           #System.OrderTable[#Chain_To_Chain_CurrentOrder].Status := #CANCELED_STATUS;
           #System.OrderTable[#Chain_To_Chain_CurrentOrder].CompleteTime := #CurrentTime;
           #Chain_To_Chain_CurrentOrder := 0;
           //#Cnv_Entry.Instruction.Execute := FALSE;
       END_IF;

       //Error
       IF (#Cnv_PopUp_2.Error OR #Cnv_PopUp_3.Error) THEN
           //#Cnv_Entry.Instruction.Execute := FALSE;
           //
           "Control_DB"."Carrousel_Order Table".Task_Data_Available := FALSE;//#System.OrderTable[#Chain_To_Chain_CurrentOrder].OPC_Control.Task_Data_Available; // Send the Task Data Available from WCS 
           "Control_DB"."Carrousel_Order Table".Task_Type := 0; //  Send the Task Type - Chain to Chain Conveyor = Task Type = 7
           "Control_DB"."Carrousel_Order Table".Task_ID := 0; // Send the Task ID number;
           "Control_DB"."Carrousel_Order Table".Task_Metadata := ''; // Send the Task Metadata Unique identifier
           "Control_DB"."Carrousel_Order Table".Source_Location := 0; // Send the Source Location from the Conveyor
           "Control_DB"."Carrousel_Order Table".Destination_Location := 0; // Send the Destination Location to the Conveyor;

           #System.OrderTable[#Chain_To_Chain_CurrentOrder].ErrorID := (#Cnv_PopUp_2.Cnv_Errors.Error_Word_1
                                                                        OR #Cnv_PopUp_3.Cnv_Errors.Error_Word_1);

       END_IF;

       //MOVEMENT FINALIZED
       #Chain_To_ChainDoneRTrig(CLK := "Control_DB"."Carrousel_Order Table".Movement_Request_Complete);
       IF #Chain_To_ChainDoneRTrig.Q THEN

           "Control_DB"."Carrousel_Order Table".Task_Data_Available := FALSE;//#System.OrderTable[#Chain_To_Chain_CurrentOrder].OPC_Control.Task_Data_Available; // Send the Task Data Available from WCS 
           "Control_DB"."Carrousel_Order Table".Task_Type := 0; //  Send the Task Type - Chain to Chain Conveyor = Task Type = 7
           "Control_DB"."Carrousel_Order Table".Task_ID := 0; // Send the Task ID number;
           "Control_DB"."Carrousel_Order Table".Task_Metadata := ''; // Send the Task Metadata Unique identifier
           "Control_DB"."Carrousel_Order Table".Source_Location := 0; // Send the Source Location from the Conveyor
           "Control_DB"."Carrousel_Order Table".Destination_Location := 0; // Send the Destination Location to the Conveyor;


           #Chain_To_Chain_WatchdogStart := FALSE;
           #System.OrderTable[#Chain_To_Chain_CurrentOrder].Status := #COMPLETED_STATUS;
           #System.OrderTable[#Chain_To_Chain_CurrentOrder].CompleteTime := #CurrentTime;
           #Chain_To_Chain_CurrentOrder := 0;
       END_IF;
   END_REGION

   REGION Pop4 to Pick Station - Carousel Conveyors - Pop 4 to Pick Station
       IF #System.OrderTable[1].StepNo <> 0
           AND #System.OrderTable[1].Device = #POP4_TO_PICK_DEVICE
           AND #System.OrderTable[1].Status = #QUEUED_STATUS
           AND NOT (#Cnv_PopUp_4.Running OR #Cnv_PopUp_1.Running)
           AND NOT #System.Error
           AND NOT #Canceling
           AND #System.OrderTable[#Roller_To_Roller_CurrentOrder].Status <> #RUNNING_STATUS
           AND #System.OrderTable[#PickSt_To_Pop1_CurrentOrder].Status <> #RUNNING_STATUS

       THEN
           #Pop4_To_PickSt_CurrentOrder := 1;
       END_IF;
       IF #System.OrderTable[#Pop4_To_PickSt_CurrentOrder].StepNo <> 0
           AND #System.OrderTable[#Pop4_To_PickSt_CurrentOrder].Device = #POP4_TO_PICK_DEVICE
           AND #System.OrderTable[#Pop4_To_PickSt_CurrentOrder].Status = #QUEUED_STATUS
           AND NOT (#Cnv_PopUp_4.Running OR #Cnv_PopUp_1.Running)
           AND NOT #System.Error
           AND NOT #Canceling
           AND #System.OrderTable[#Roller_To_Roller_CurrentOrder].Status <> #RUNNING_STATUS
           AND #System.OrderTable[#PickSt_To_Pop1_CurrentOrder].Status <> #RUNNING_STATUS
       THEN
           //OPC Commands to Move Pallets - Carousel Conveyors
           // WCS => Order Table => OPC Ua Control Table

           "Control_DB"."Carrousel_Order Table".Task_Data_Available := TRUE;//#System.OrderTable[#Pop4_To_PickSt_CurrentOrder].OPC_Control.Task_Data_Available; // Send the Task Data Available from WCS 
           "Control_DB"."Carrousel_Order Table".Task_Type := #System.OrderTable[#Pop4_To_PickSt_CurrentOrder].OPC_Control.Task_Type; //  Send the Task Type - Pop4 to Pick Station Conveyor = Task Type = 8
           "Control_DB"."Carrousel_Order Table".Task_ID := #System.OrderTable[#Pop4_To_PickSt_CurrentOrder].OPC_Control.Task_ID; // Send the Task ID number;
           "Control_DB"."Carrousel_Order Table".Task_Metadata := #System.OrderTable[#Pop4_To_PickSt_CurrentOrder].OPC_Control.Task_Metadata; // Send the Task Metadata Unique identifier
           "Control_DB"."Carrousel_Order Table".Source_Location := #System.OrderTable[#Pop4_To_PickSt_CurrentOrder].OPC_Control.Source_Location; // Send the Source Location from the Conveyor
           "Control_DB"."Carrousel_Order Table".Destination_Location := #System.OrderTable[#Pop4_To_PickSt_CurrentOrder].OPC_Control.Destination_Location; // Send the Destination Location to the Conveyor;
           #Pop4_To_PickWatchdogStart := TRUE;



       END_IF;

       //RUNNING
       IF (#Cnv_PopUp_4.Running OR #Cnv_PopUp_1.Running) AND #System.Auto_Man THEN
           //#Cnv_Entry.Instruction.Execute := FALSE;
           #System.OrderTable[#Pop4_To_PickSt_CurrentOrder].Status := #RUNNING_STATUS;
       END_IF;

       //Cancel order
       IF #Canceling AND NOT (#Cnv_PopUp_4.Running OR #Cnv_PopUp_1.Running) AND #Pop4_To_PickSt_CurrentOrder <> 0 THEN
           #System.OrderTable[#Pop4_To_PickSt_CurrentOrder].Status := #CANCELED_STATUS;
           #System.OrderTable[#Pop4_To_PickSt_CurrentOrder].CompleteTime := #CurrentTime;
           #Pop4_To_PickSt_CurrentOrder := 0;

           "Control_DB"."Carrousel_Order Table".Task_Data_Available := FALSE;//#System.OrderTable[#Chain_To_Chain_CurrentOrder].OPC_Control.Task_Data_Available; // Send the Task Data Available from WCS 
           "Control_DB"."Carrousel_Order Table".Task_Type := 0; //  Send the Task Type - Chain to Chain Conveyor = Task Type = 7
           "Control_DB"."Carrousel_Order Table".Task_ID := 0; // Send the Task ID number;
           "Control_DB"."Carrousel_Order Table".Task_Metadata := ''; // Send the Task Metadata Unique identifier
           "Control_DB"."Carrousel_Order Table".Source_Location := 0; // Send the Source Location from the Conveyor
           "Control_DB"."Carrousel_Order Table".Destination_Location := 0; // Send the Destination Location to the Conveyor;

           //#Cnv_Entry.Instruction.Execute := FALSE;
       END_IF;

       //Error
       IF (#Cnv_PopUp_4.Error OR #Cnv_PopUp_1.Error) THEN
           //#Cnv_Entry.Instruction.Execute := FALSE;
           "Control_DB"."Carrousel_Order Table".Task_Data_Available := FALSE;//#System.OrderTable[#Chain_To_Chain_CurrentOrder].OPC_Control.Task_Data_Available; // Send the Task Data Available from WCS 
           "Control_DB"."Carrousel_Order Table".Task_Type := 0; //  Send the Task Type - Chain to Chain Conveyor = Task Type = 7
           "Control_DB"."Carrousel_Order Table".Task_ID := 0; // Send the Task ID number;
           "Control_DB"."Carrousel_Order Table".Task_Metadata := ''; // Send the Task Metadata Unique identifier
           "Control_DB"."Carrousel_Order Table".Source_Location := 0; // Send the Source Location from the Conveyor
           "Control_DB"."Carrousel_Order Table".Destination_Location := 0; // Send the Destination Location to the Conveyor;
           #System.OrderTable[#Pop4_To_PickSt_CurrentOrder].ErrorID := (#Cnv_PopUp_4.Cnv_Errors.Error_Word_1
           OR #Cnv_PopUp_1.Cnv_Errors.Error_Word_1);

       END_IF;

       //MOVEMENT FINALIZED
       #Pop4_To_PickSt_DoneRTrig(CLK := "Control_DB"."Carrousel_Order Table".Movement_Request_Complete);
       IF #Pop4_To_PickSt_DoneRTrig.Q THEN
           #Pop4_To_PickWatchdogStart := FALSE;

           "Control_DB"."Carrousel_Order Table".Task_Data_Available := FALSE;//#System.OrderTable[#Chain_To_Chain_CurrentOrder].OPC_Control.Task_Data_Available; // Send the Task Data Available from WCS 
           "Control_DB"."Carrousel_Order Table".Task_Type := 0; //  Send the Task Type - Chain to Chain Conveyor = Task Type = 7
           "Control_DB"."Carrousel_Order Table".Task_ID := 0; // Send the Task ID number;
           "Control_DB"."Carrousel_Order Table".Task_Metadata := ''; // Send the Task Metadata Unique identifier
           "Control_DB"."Carrousel_Order Table".Source_Location := 0; // Send the Source Location from the Conveyor
           "Control_DB"."Carrousel_Order Table".Destination_Location := 0; // Send the Destination Location to the Conveyor;

           #System.OrderTable[#Pop4_To_PickSt_CurrentOrder].Status := #COMPLETED_STATUS;
           #System.OrderTable[#Pop4_To_PickSt_CurrentOrder].CompleteTime := #CurrentTime;
           #Pop4_To_PickSt_CurrentOrder := 0;
       END_IF;
   END_REGION

   REGION Pick Station to Pop1 - Carousel Conveyors - Pick Station To Pop 1 
       IF #System.OrderTable[1].StepNo <> 0
           AND #System.OrderTable[1].Device = #PICK_TO_POP1_DEVICE
           AND #System.OrderTable[1].Status = #QUEUED_STATUS
           AND NOT (#Cnv_PopUp_1.Running)
           AND NOT #System.Error
           AND NOT #Canceling
           AND #System.OrderTable[#Roller_To_Roller_CurrentOrder].Status <> #RUNNING_STATUS
           AND #System.OrderTable[#Pop4_To_PickSt_CurrentOrder].Status <> #RUNNING_STATUS
       THEN
           #PickSt_To_Pop1_CurrentOrder := 1;
       END_IF;
       IF #System.OrderTable[#PickSt_To_Pop1_CurrentOrder].StepNo <> 0
           AND #System.OrderTable[#PickSt_To_Pop1_CurrentOrder].Device = #PICK_TO_POP1_DEVICE
           AND #System.OrderTable[#PickSt_To_Pop1_CurrentOrder].Status = #QUEUED_STATUS
           AND NOT (#Cnv_PopUp_1.Running)
           AND NOT #System.Error
           AND NOT #Canceling
           AND #System.OrderTable[#Roller_To_Roller_CurrentOrder].Status <> #RUNNING_STATUS
           AND #System.OrderTable[#Pop4_To_PickSt_CurrentOrder].Status <> #RUNNING_STATUS
       THEN
           //OPC Commands to Move Pallets - Carousel Conveyors
           // WCS => Order Table => OPC Ua Control Table

           "Control_DB"."Carrousel_Order Table".Task_Data_Available := TRUE;//#System.OrderTable[#PickSt_To_Pop1_CurrentOrder].OPC_Control.Task_Data_Available; // Send the Task Data Available from WCS 
           "Control_DB"."Carrousel_Order Table".Task_Type := #System.OrderTable[#PickSt_To_Pop1_CurrentOrder].OPC_Control.Task_Type; //  Send the Task Type - Roller to Roller Conveyor = Task Type = 6
           "Control_DB"."Carrousel_Order Table".Task_ID := #System.OrderTable[#PickSt_To_Pop1_CurrentOrder].OPC_Control.Task_ID; // Send the Task ID number;
           "Control_DB"."Carrousel_Order Table".Task_Metadata := #System.OrderTable[#PickSt_To_Pop1_CurrentOrder].OPC_Control.Task_Metadata; // Send the Task Metadata Unique identifier
           "Control_DB"."Carrousel_Order Table".Source_Location := #System.OrderTable[#PickSt_To_Pop1_CurrentOrder].OPC_Control.Source_Location; // Send the Source Location from the Conveyor
           "Control_DB"."Carrousel_Order Table".Destination_Location := #System.OrderTable[#PickSt_To_Pop1_CurrentOrder].OPC_Control.Destination_Location; // Send the Destination Location to the Conveyor;
           #PickSt_To_Pop1WatchdogStart := true;


       END_IF;

       //RUNNING
       IF (#Cnv_PopUp_1.Running) AND #System.Auto_Man THEN
           //#Cnv_Entry.Instruction.Execute := FALSE;
           #System.OrderTable[#PickSt_To_Pop1_CurrentOrder].Status := #RUNNING_STATUS;
       END_IF;

       //Cancel order
       IF #Canceling AND NOT (#Cnv_PopUp_1.Running) AND #PickSt_To_Pop1_CurrentOrder <> 0 THEN
           #System.OrderTable[#PickSt_To_Pop1_CurrentOrder].Status := #CANCELED_STATUS;
           #System.OrderTable[#PickSt_To_Pop1_CurrentOrder].CompleteTime := #CurrentTime;
           #PickSt_To_Pop1_CurrentOrder := 0;
           "Control_DB"."Carrousel_Order Table".Task_Data_Available := FALSE;//#System.OrderTable[#Chain_To_Chain_CurrentOrder].OPC_Control.Task_Data_Available; // Send the Task Data Available from WCS 
           "Control_DB"."Carrousel_Order Table".Task_Type := 0; //  Send the Task Type - Chain to Chain Conveyor = Task Type = 7
           "Control_DB"."Carrousel_Order Table".Task_ID := 0; // Send the Task ID number;
           "Control_DB"."Carrousel_Order Table".Task_Metadata := ''; // Send the Task Metadata Unique identifier
           "Control_DB"."Carrousel_Order Table".Source_Location := 0; // Send the Source Location from the Conveyor
           "Control_DB"."Carrousel_Order Table".Destination_Location := 0; // Send the Destination Location to the Conveyor;
           //#Cnv_Entry.Instruction.Execute := FALSE;
       END_IF;

       //Error
       IF (#Cnv_PopUp_2.Error OR #Cnv_PopUp_3.Error) THEN
           //#Cnv_Entry.Instruction.Execute := FALSE;
           "Control_DB"."Carrousel_Order Table".Task_Data_Available := FALSE;//#System.OrderTable[#Chain_To_Chain_CurrentOrder].OPC_Control.Task_Data_Available; // Send the Task Data Available from WCS 
           "Control_DB"."Carrousel_Order Table".Task_Type := 0; //  Send the Task Type - Chain to Chain Conveyor = Task Type = 7
           "Control_DB"."Carrousel_Order Table".Task_ID := 0; // Send the Task ID number;
           "Control_DB"."Carrousel_Order Table".Task_Metadata := ''; // Send the Task Metadata Unique identifier
           "Control_DB"."Carrousel_Order Table".Source_Location := 0; // Send the Source Location from the Conveyor
           "Control_DB"."Carrousel_Order Table".Destination_Location := 0; // Send the Destination Location to the Conveyor;
           #System.OrderTable[#PickSt_To_Pop1_CurrentOrder].ErrorID := (#Cnv_PopUp_2.Cnv_Errors.Error_Word_1
           OR #Cnv_PopUp_3.Cnv_Errors.Error_Word_1);

       END_IF;

       //MOVEMENT FINALIZED
       #PickSt_To_Pop1_DoneRTrig(CLK := "Control_DB"."Carrousel_Order Table".Movement_Request_Complete);
       IF #PickSt_To_Pop1_DoneRTrig.Q THEN

           "Control_DB"."Carrousel_Order Table".Task_Data_Available := FALSE;//#System.OrderTable[#Chain_To_Chain_CurrentOrder].OPC_Control.Task_Data_Available; // Send the Task Data Available from WCS 
           "Control_DB"."Carrousel_Order Table".Task_Type := 0; //  Send the Task Type - Chain to Chain Conveyor = Task Type = 7
           "Control_DB"."Carrousel_Order Table".Task_ID := 0; // Send the Task ID number;
           "Control_DB"."Carrousel_Order Table".Task_Metadata := ''; // Send the Task Metadata Unique identifier
           "Control_DB"."Carrousel_Order Table".Source_Location := 0; // Send the Source Location from the Conveyor
           "Control_DB"."Carrousel_Order Table".Destination_Location := 0; // Send the Destination Location to the Conveyor;

           #PickSt_To_Pop1WatchdogStart := FALSE;
           #System.OrderTable[#PickSt_To_Pop1_CurrentOrder].Status := #COMPLETED_STATUS;
           #System.OrderTable[#PickSt_To_Pop1_CurrentOrder].CompleteTime := #CurrentTime;
           #PickSt_To_Pop1_CurrentOrder := 0;
       END_IF;
   END_REGION

   REGION Weigh Station - Carousel Conveyors 
       IF #System.OrderTable[1].StepNo <> 0
           AND #System.OrderTable[1].Device = #WEIGH_STATION_DEVICE
           AND #System.OrderTable[1].Status = #QUEUED_STATUS
           AND NOT ("Control_DB"."Weighing Station".Running)
           AND NOT #System.Error
           AND NOT #Canceling
       THEN
           #WeighingStation_CurrentOrder := 1;
       END_IF;
       IF #System.OrderTable[#WeighingStation_CurrentOrder].StepNo <> 0
           AND #System.OrderTable[#WeighingStation_CurrentOrder].Device = #WEIGH_STATION_DEVICE
           AND #System.OrderTable[#WeighingStation_CurrentOrder].Status = #QUEUED_STATUS
           AND NOT ("Control_DB"."Weighing Station".Running)
           AND NOT #System.Error
           AND NOT #Canceling
       THEN
           //OPC Commands to Move Pallets - Carousel Conveyors
           // WCS => Order Table => OPC Ua Control Table


           "Control_DB"."Carrousel_Order Table".Task_Data_Available := TRUE;//#System.OrderTable[#WeighingStation_CurrentOrder].OPC_Control.Task_Data_Available; // Send the Task Data Available from WCS 
           "Control_DB"."Carrousel_Order Table".Task_Type := #System.OrderTable[#WeighingStation_CurrentOrder].OPC_Control.Task_Type; //  Send the Task Type - Start Weigh Station = Task Type = 10
           "Control_DB"."Carrousel_Order Table".Task_ID := #System.OrderTable[#WeighingStation_CurrentOrder].OPC_Control.Task_ID; // Send the Task ID number;
           "Control_DB"."Carrousel_Order Table".Task_Metadata := #System.OrderTable[#WeighingStation_CurrentOrder].OPC_Control.Task_Metadata; // Send the Task Metadata Unique identifier
           #WeighingStation_WatchdogStart := true;


       END_IF;

       //RUNNING
       IF ("Control_DB"."Weighing Station".Running) AND #System.Auto_Man THEN
           //#Cnv_Entry.Instruction.Execute := FALSE;
           #System.OrderTable[#WeighingStation_CurrentOrder].Status := #RUNNING_STATUS;

       END_IF;

       //Cancel order
       IF #Canceling AND NOT ("Control_DB"."Weighing Station".Running) AND #WeighingStation_CurrentOrder <> 0 THEN
           #System.OrderTable[#WeighingStation_CurrentOrder].Status := #CANCELED_STATUS;
           #System.OrderTable[#WeighingStation_CurrentOrder].CompleteTime := #CurrentTime;
           #WeighingStation_CurrentOrder := 0;
           //#Cnv_Entry.Instruction.Execute := FALSE;
           "Control_DB"."Carrousel_Order Table".Task_Data_Available := FALSE;//#System.OrderTable[#WeighingStation_CurrentOrder].OPC_Control.Task_Data_Available; // Send the Task Data Available from WCS 
           "Control_DB"."Carrousel_Order Table".Task_Type := 0; //  Send the Task Type - Start Weigh Station = Task Type = 10
           "Control_DB"."Carrousel_Order Table".Task_ID := 0; // Send the Task ID number;
           "Control_DB"."Carrousel_Order Table".Task_Metadata := ''; // Send the Task Metadata Unique identifier
       END_IF;
     (*  
       //Error
       IF (#WeighingStation. OR #Cnv_PopUp_3.Error) THEN
           //#Cnv_Entry.Instruction.Execute := FALSE;

           #System.OrderTable[#WeighingStation_CurrentOrder].ErrorID := (#Cnv_PopUp_2.Cnv_Errors.Error_Word_1
         OR #Cnv_PopUp_3.Cnv_Errors.Error_Word_1);

       END_IF;
      *) 
       //MOVEMENT FINALIZED
       #WeighingStationDoneRTrig(CLK := "Control_DB"."Weighing Station".Done);
       IF #WeighingStationDoneRTrig.Q THEN
           #WeighingStation_WatchdogStart := FALSE;
           #System.OrderTable[#WeighingStation_CurrentOrder].Status := #COMPLETED_STATUS;
           #System.OrderTable[#WeighingStation_CurrentOrder].CompleteTime := #CurrentTime;
           #WeighingStation_CurrentOrder := 0;

           "Control_DB"."Carrousel_Order Table".Task_Data_Available := FALSE;//#System.OrderTable[#WeighingStation_CurrentOrder].OPC_Control.Task_Data_Available; // Send the Task Data Available from WCS 
           "Control_DB"."Carrousel_Order Table".Task_Type := 0; //  Send the Task Type - Start Weigh Station = Task Type = 10
           "Control_DB"."Carrousel_Order Table".Task_ID := 0; // Send the Task ID number;
           "Control_DB"."Carrousel_Order Table".Task_Metadata := ''; // Send the Task Metadata Unique identifier
       END_IF;
   END_REGION
   (*
   REGION Profile Station - Carousel Conveyors 
       IF #System.OrderTable[1].StepNo <> 0
           AND #System.OrderTable[1].Device = #PROFILE_STATION_DEVICE
           AND #System.OrderTable[1].Status = #QUEUED_STATUS
           AND NOT ("Control_DB"."Profiling Station".Running)
           AND NOT #System.Error
           AND NOT #Canceling
       THEN
           #ProfileStation_CurrentOrder := 1;
       END_IF;
       IF #System.OrderTable[#ProfileStation_CurrentOrder].StepNo <> 0
           AND #System.OrderTable[#ProfileStation_CurrentOrder].Device = #PROFILE_STATION_DEVICE
           AND #System.OrderTable[#ProfileStation_CurrentOrder].Status = #QUEUED_STATUS
           AND NOT ("Control_DB"."Profiling Station".Running)
           AND NOT #System.Error
           AND NOT #Canceling
       THEN
           //OPC Commands to Move Pallets - Carousel Conveyors
           // WCS => Order Table => OPC Ua Control Table

           "Control_DB"."Carrousel_Order Table".Task_Data_Available := TRUE;//#System.OrderTable[#ProfileStation_CurrentOrder].OPC_Control.Task_Data_Available; // Send the Task Data Available from WCS 
           "Control_DB"."Carrousel_Order Table".Task_Type := #System.OrderTable[#ProfileStation_CurrentOrder].OPC_Control.Task_Type; //  Send the Task Type - Start Weigh Station = Task Type = 10
           "Control_DB"."Carrousel_Order Table".Task_ID := #System.OrderTable[#ProfileStation_CurrentOrder].OPC_Control.Task_ID; // Send the Task ID number;
           "Control_DB"."Carrousel_Order Table".Task_Metadata := #System.OrderTable[#ProfileStation_CurrentOrder].OPC_Control.Task_Metadata; // Send the Task Metadata Unique identifier
           #ProfileStation_WatchdogStart := true;


       END_IF;

       //RUNNING
       IF ("Control_DB"."Profiling Station".Running) AND #System.Auto_Man THEN
           //#Cnv_Entry.Instruction.Execute := FALSE;
           #System.OrderTable[#ProfileStation_CurrentOrder].Status := #RUNNING_STATUS;

           "Control_DB"."Carrousel_Order Table".Task_Data_Available := FALSE;//#System.OrderTable[#ProfileStation_CurrentOrder].OPC_Control.Task_Data_Available; // Send the Task Data Available from WCS 
           "Control_DB"."Carrousel_Order Table".Task_Type := 0; //  Send the Task Type - Start Weigh Station = Task Type = 10
           "Control_DB"."Carrousel_Order Table".Task_ID := 0; // Send the Task ID number;
           "Control_DB"."Carrousel_Order Table".Task_Metadata := ''; // Send the Task Metadata Unique identifier
           #ProfileStation_WatchdogStart := true;
       END_IF;

       //Cancel order
       IF #Canceling AND NOT ("Control_DB"."Profiling Station".Running) AND #ProfileStation_CurrentOrder <> 0 THEN
           #System.OrderTable[#ProfileStation_CurrentOrder].Status := #CANCELED_STATUS;
           #System.OrderTable[#ProfileStation_CurrentOrder].CompleteTime := #CurrentTime;
           #ProfileStation_CurrentOrder := 0;
           "Control_DB"."Carrousel_Order Table".Task_Data_Available := FALSE;//#System.OrderTable[#ProfileStation_CurrentOrder].OPC_Control.Task_Data_Available; // Send the Task Data Available from WCS 
           "Control_DB"."Carrousel_Order Table".Task_Type := 0; //  Send the Task Type - Start Weigh Station = Task Type = 10
           "Control_DB"."Carrousel_Order Table".Task_ID := 0; // Send the Task ID number;
           "Control_DB"."Carrousel_Order Table".Task_Metadata := ''; // Send the Task Metadata Unique identifier
           //#Cnv_Entry.Instruction.Execute := FALSE;
       END_IF;
       (*  
         //Error
         IF (#WeighingStation. OR #Cnv_PopUp_3.Error) THEN
             //#Cnv_Entry.Instruction.Execute := FALSE;

             #System.OrderTable[#WeighingStation_CurrentOrder].ErrorID := (#Cnv_PopUp_2.Cnv_Errors.Error_Word_1
           OR #Cnv_PopUp_3.Cnv_Errors.Error_Word_1);

         END_IF;
        *)
        //MOVEMENT FINALIZED
       #ProfileStationDoneRTrig(CLK := "Control_DB"."Profiling Station".Done);
       IF #ProfileStationDoneRTrig.Q THEN
            #ProfileStation_WatchdogStart := FALSE;
            #System.OrderTable[#ProfileStation_CurrentOrder].Status := #COMPLETED_STATUS;
            #System.OrderTable[#ProfileStation_CurrentOrder].CompleteTime := #CurrentTime;
            #ProfileStation_CurrentOrder := 0;
            "Control_DB"."Carrousel_Order Table".Task_Data_Available := FALSE;//#System.OrderTable[#ProfileStation_CurrentOrder].OPC_Control.Task_Data_Available; // Send the Task Data Available from WCS 
            "Control_DB"."Carrousel_Order Table".Task_Type := 0; //  Send the Task Type - Start Weigh Station = Task Type = 10
            "Control_DB"."Carrousel_Order Table".Task_ID := 0; // Send the Task ID number;
            "Control_DB"."Carrousel_Order Table".Task_Metadata := ''; // Send the Task Metadata Unique identifier
        END_IF;
    END_REGION
   *)
   REGION Max Running Order Number
       #MaxRunningOrderNo := MAX(IN1 := #Roller_To_Roller_CurrentOrder, IN2 := #Chain_To_Chain_CurrentOrder,
                                 IN3 := #Pop4_To_PickSt_CurrentOrder, IN4 := #PickSt_To_Pop1_CurrentOrder,
                                 IN5 := #WeighingStation_CurrentOrder, IN6 := #ProfileStation_CurrentOrder);
   END_REGION

   REGION Pause Orders
       #ErrorRTrig(CLK := #System.Error);
       #PauseRTrig(CLK := #System.PauseOrders OR NOT #System.Auto_Man);
       IF #ErrorRTrig.Q OR #PauseRTrig.Q THEN
           #System.PauseOrders := FALSE;
           #System.Paused := #MaxRunningOrderNo > 0;
           IF #System.Paused THEN
               FOR #i := 1 TO UDINT_TO_DINT(#MaxRunningOrderNo) DO
                   IF #System.OrderTable[#i].Status = '' THEN
                       EXIT;
                   ELSIF #System.OrderTable[#i].Status = #QUEUED_STATUS THEN
                       #System.OrderTable[#i].Status := #PAUSED_STATUS;
                   ELSIF #System.OrderTable[#i].Status = #RUNNING_STATUS AND NOT #System.Auto_Man THEN
                       #System.OrderTable[#i].Status := #CANCELED_STATUS;
                   END_IF;
               END_FOR;
           END_IF;
       END_IF;
       IF #System.Paused AND #MaxRunningOrderNo = 0 THEN
           #System.Paused := FALSE;
       END_IF;
   END_REGION

   REGION Cancel Orders
       #CancelRTrig(CLK := #System.CancelOrders);
       #WeighingStation.Cancel := #ProfileStation.Cancel := #CancelRTrig.Q;
       IF #CancelRTrig.Q THEN
           #Canceling := TRUE;
           #System.CancelOrders := FALSE;
           #System.Paused := FALSE;
           FOR #i := 1 TO UDINT_TO_DINT(#MaxRunningOrderNo) DO
               IF #System.OrderTable[#i].Status = '' THEN
                   CONTINUE;
               ELSIF #System.OrderTable[#i].Status = #PAUSED_STATUS
                   OR #System.OrderTable[#i].Status = #QUEUED_STATUS
               THEN
                   #System.OrderTable[#i].Status := #CANCELED_STATUS;
                   #System.OrderTable[#i].CompleteTime := #CurrentTime;
               ELSIF #System.OrderTable[#i].Status = #ERROR_STATUS
               THEN
                   #System.OrderTable[#i].Status := #ERROR_CANCELED_STATUS;
                   #System.OrderTable[#i].CompleteTime := #CurrentTime;
               END_IF;
           END_FOR;
           #System.CurrentOrder := 0;
       END_IF;
       IF #Canceling AND NOT (#Cnv_Entry.Running OR #Cnv_PopUp_1.Running OR #WeighingStation.Running OR #ProfileStation.Running
           OR #Cnv_PopUp_2.Running OR #Cnv_PopUp_3.Running OR #Cnv_PopUp_4.Running OR #Cnv_Exit.Running) THEN
           #Canceling := FALSE;
           #Roller_To_Roller_CurrentOrder := #Chain_To_Chain_CurrentOrder:= #PickSt_To_Pop1_CurrentOrder := #Pop4_To_PickSt_CurrentOrder := 0;
            #WeighingStation_CurrentOrder:= #ProfileStation_CurrentOrder := 0;
       END_IF;
   END_REGION

   REGION Resume Orders
       #ResumeRTrig(CLK := #System.ResumeOrders);
       IF #ResumeRTrig.Q THEN
           #System.ResumeOrders := FALSE;
           #System.CurrentOrder := #MaxRunningOrderNo;
           IF NOT #System.Error THEN
               #System.Paused := FALSE;
               FOR #i := 1 TO UDINT_TO_DINT(#MaxRunningOrderNo) DO
                   IF #System.OrderTable[#i].Status = '' THEN
                       EXIT;
                   ELSIF #System.OrderTable[#i].Status = #PAUSED_STATUS
                       OR #System.OrderTable[#i].Status = #ERROR_STATUS
                   THEN
                       #System.OrderTable[#i].Status := #QUEUED_STATUS;
                   END_IF;
               END_FOR;
           END_IF;

       END_IF;
   END_REGION

   REGION Order Handler
       IF #System.Running AND NOT #System.Error
           AND (#System.OrderTable[#System.CurrentOrder].Status = #COMPLETED_STATUS
           OR #System.OrderTable[#System.CurrentOrder].Status = #ERROR_STATUS
           OR #System.OrderTable[#System.CurrentOrder].Status = #ERROR_CANCELED_STATUS
           OR #System.OrderTable[#System.CurrentOrder].Sequence = 0)
       THEN
           IF #System.CurrentOrder > 0 THEN
               #System.CurrentOrder -= 1;
           ELSE
               #System.CurrentOrder := 0;
           END_IF;
       END_IF;
   END_REGION

   REGION Watchdogs
       //Watchdog Timers
       #PickSt_To_Pop1WatchdogTimer(IN := #PickSt_To_Pop1WatchdogStart,
                                    PT := UDINT_TO_TIME(#Watchdog.Pick_TO_Pop1 * 60000),
                                    Q => #System.Watchdog_TimeOut.Pick_TO_Pop1);
       #Roller_To_Roller_WatchdogTimer(IN := #Roller_To_Roller_WatchdogStart,
                                       PT := UDINT_TO_TIME(#Watchdog.Roller_TO_Roller * 60000),
                                       Q => #System.Watchdog_TimeOut.Roller_TO_Roller);
       #Chain_To_Chain_WatchdogTimer(IN := #Chain_To_Chain_WatchdogStart,
                                     PT := UDINT_TO_TIME(#Watchdog.Chain_TO_Chain * 60000),
                                     Q => #System.Watchdog_TimeOut.Chain_TO_Chain);
       #Pop4_To_PickWatchdogTimer(IN := #Pop4_To_PickWatchdogStart,
                                  PT := UDINT_TO_TIME(#Watchdog.Pop4_TO_Pick * 60000),
                                  Q => #System.Watchdog_TimeOut.Pop4_TO_Pick);
       #WeighingStation_WatchdogTimer(IN := #WeighingStation_WatchdogStart,
                                      PT := UDINT_TO_TIME(#Watchdog.Weigh_Station * 60000),
                                      Q => #System.Watchdog_TimeOut.Weigh_Station);
       #ProfileStation_WatchdogTimer(IN := #ProfileStation_WatchdogStart,
                                     PT := UDINT_TO_TIME(#Watchdog.Profile_Station * 60000),
                                     Q => #System.Watchdog_TimeOut.Profile_Station);

       //Reset  Watchdog Timers
       IF #System.Error OR #CancelRTrig.Q OR #PauseRTrig.Q OR "Reset_All" THEN
           #PickSt_To_Pop1WatchdogStart := FALSE;
           #Roller_To_Roller_WatchdogStart := FALSE;
           #Chain_To_Chain_WatchdogStart := FALSE;
           #Pop4_To_PickWatchdogStart := FALSE;
           #WeighingStation_WatchdogStart := FALSE;
           #ProfileStation_WatchdogStart := FALSE;

       END_IF;
   END_REGION

   REGION Reset Next Order Number
       IF #System.NextOrder > 1
           AND #CurrentDTL.HOUR = 0
           AND #CurrentDTL.MINUTE = 0
           AND #CurrentDTL.SECOND = 0
       THEN
           #System.NextOrder := 1;
       END_IF;

   END_REGION

   REGION #System Mode and State
       #System.Selected := #System_Selected; // System selected
       #System.Ready := NOT #System.Error AND #System.Selected;
       #System.Auto_Man := #AutoMan_Switch;
       #System.Running := #Cnv_Entry.Running OR #Cnv_PopUp_1.Running OR #WeighingStation.Running
       OR #ProfileStation.Running OR #Cnv_PopUp_3.Running OR #Cnv_PopUp_4.Running;

       #System.Error := #Cnv_Entry.Error OR #Cnv_PopUp_1.Error OR #Cnv_PopUp_2.Error OR #Cnv_PopUp_3.Error OR #Cnv_PopUp_4.Error
       OR #Cnv_Exit.Error ; (*Implement Weigh station error and Profile Station error*)
       #System.IDLE := NOT #System.Running AND NOT #System.Paused AND NOT #System.Error;
       IF #System.Running THEN
           #System.State := 1;
       ELSIF #System.Paused AND NOT #System.Error THEN
           #System.State := 2;
       ELSIF #System.Error THEN
           #System.State := 3;
       ELSE
           #System.State := 0;
       END_IF;
   END_REGION
END_FUNCTION_BLOCK

FUNCTION_BLOCK "PConveyor_1_FB_1"   // FB36, SCL
TITLE = Conveyor Instance FB
{ S7_Optimized_Access := 'TRUE' }
AUTHOR : Mertin Coetzee
VERSION : 0.1
// stored: AutoNumber true, IsIECCheckEnabled false, IsRetainMemResEnabled false, MemoryReserve 100, SetENOAutomatically false, UDAEnableTagReadback false
   VAR_INPUT
      Cnv_Settings : "PopUp_Cnv_Settings";
   END_VAR
   VAR_IN_OUT
      Cnv_Control : "PopUp_Cnv_Control";
      SinaSpeed_Roller : SinaSpeed;
      SinaSpeed_Chain : SinaSpeed;
      SinaSpeed_Lift : SinaSpeed;
   END_VAR
   VAR
      State : UInt;
      Timer_TC : TON_TIME;
      Timer_Transfer { S7_SetPoint := 'True'} : TON_TIME;
      Watchdog { S7_SetPoint := 'True'} : TON_TIME;
      Transfer_Direction { S7_SetPoint := 'True'} : String;
      MainSetpoint_Roller : Int;
      MainSetpoint_Chain : Int;
      MainSetpoint_Lift : Int;
      IEC_Timer_0_Instance_1 { S7_SetPoint := 'True'} : TON_TIME;
      R_TRIG_Instance { S7_SetPoint := 'True'} : R_TRIG;
   END_VAR
   VAR_TEMP
      Execute_Old : Bool;
      Stop_Old : Bool;
   END_VAR
BEGIN
   "R_TRIG_DB_13"(CLK := #Cnv_Control.Instruction.Execute AND NOT #Execute_Old);
   "R_TRIG_DB_14"(CLK := #Cnv_Control.Instruction.Stop AND NOT #Stop_Old);

   #Execute_Old := #Cnv_Control.Instruction.Execute;
   #Stop_Old := #Cnv_Control.Instruction.Stop;

   #Cnv_Control.Enabled := #Cnv_Control.Instruction.Enable;

   //MODES
   #Cnv_Control.Mode := #Cnv_Control.Instruction.Mode_Change;
   IF (#Cnv_Control.Mode = 1 OR #Cnv_Control.Mode = 5) AND NOT #Cnv_Control.Error THEN
       #State := 500;
   END_IF;

   #R_TRIG_Instance(CLK := #Cnv_Control.Mode = 3);
   IF #R_TRIG_Instance.Q THEN
       #State := 0;
   END_IF;

   (*
   TODO:
   01. Need to add statemachine watchdog - Done
   02. Extractor needs to be on same floor for pallet to be moved in manual passed Rbwd - Done
   03. Complete reset state - Done
   04. Add stop inputs - Done
   05. Need to add variable motor speed, manual needs to be slower. - Done
   06. Need to add cyclic error checking. For odd sensor combinations as well - Partially done
   07. Need to add Shuttle monitor - Done
   08. Need to add Task ID check and start bit check to outbound pallet move. Check direction of pallet movement based on connected Cnv.
   09. Need to add checks for wrong direction of travel - Done
   10. Add checks for unsafe conditions with Cnv_Inputs - Partially Done
   11. Define Error codes - DOne
   12. Add watchdof time to Cnv Settings - Done
   13. Add self-timeout on manual 
   14. For shuttle in place sensor checks take into account extractor floor and safety stopper state
   15. Confirm modes and states are correct (Semi-auto and maintenance as well)
   16. Add the correct transfer process for the logistex-spacemaker pallet handovers.

   Mode select is done via the HMI. Might add external mode select switches.

           Mode select mask:
           0: Disabled
           1: Manual
           2: Semi-Auto
           3: Auto
           4: Teach - N/A for Cnv
           5: Maintenance

   Device ID Format: XXYYZZ    
   XX = Device type   
       01   VTD
       10  Cnv_Front_of_VTD
       11  Cnv_Rear_of_VTD
       12  Cnv_On_Extractor
       20  Safety_Stop_Front_of_VTD
       21  Safety_Stop_Rear_of_VTD
   YY = Floor   
   ZZ = VTD Connected to    
   Example: 110203 Conveyor at the rear of VTD 3 on level 2

   Pallet Alignment
   0 = no alignment
   1 = center alignment
   2 = Left
   3 = Right

    Sensor order for the conveyor:
    Lfwd Lpd1 Lpd2
     []   []   []
    ##############################
    #        Pallet Flow         #
    #         ------->>          #
    #                            #
    #                            #
    ##############################
                     []   []   []
                    Rpd2 Rpd1 Rbwd      
   *)

   REGION Cyclic Checks    
       // Update the pallet type as the Cnv_Inputs are triggered.
       #Cnv_Control.Cnv_Occupied := "PopUp Conveyor 2 - Pallet present 3";

       // Update the Cnv_Control opbject
       #Cnv_Control.SM_State := #State;
       #Cnv_Control.Stopped := NOT #Cnv_Control.Running;
       IF #Cnv_Control.Instruction.Inbound_Ready OR #Cnv_Control.Instruction.Outbound_Ready THEN
           #Cnv_Control.Ready_For_Task := TRUE;
       ELSE
           #Cnv_Control.Ready_For_Task := FALSE;
       END_IF;
   END_REGION

   REGION Auto/Semi auto mode
       CASE #State OF
           0: //Initialization
               #Cnv_Control.Instruction.Transfer_Complete := 0;
               #Cnv_Control.Instruction.Transfer_in_Progress := FALSE;
               #Cnv_Control.Running := FALSE;
               #Cnv_Control.Roller_Motor.Forward := FALSE;
               #Cnv_Control.Roller_Motor.Reverse := FALSE;
               #Cnv_Control.Roller_Motor.Speed := 0;
               #Cnv_Control.Chain_Motor.Forward := FALSE;
               #Cnv_Control.Chain_Motor.Reverse := FALSE;
               #Cnv_Control.Chain_Motor.Speed := 0;
               #Cnv_Control.Lift_Motor.Forward := FALSE;
               #Cnv_Control.Lift_Motor.Reverse := FALSE;
               #Cnv_Control.Lift_Motor.Speed := 0;
               #Transfer_Direction := '';
               #Timer_Transfer(IN := FALSE,
                               PT := T#0ms);
               IF #Cnv_Control.Enabled AND (#Cnv_Control.Mode = 3 OR #Cnv_Control.Mode = 2) AND #Cnv_Control.Error = 0 THEN
                   #State := 10;
               END_IF;

           10: //Standby - Conveyor ready to receive instruction
               IF ("R_TRIG_DB_13".Q OR #Cnv_Control.Instruction.Start_Transfer) THEN
                   //Inbound Transfer
                   IF #Cnv_Control.Instruction.Inbound_Ready AND NOT #Cnv_Control.Running AND #Cnv_Control.Error = 0 THEN
                       //Check transfer ID FROM Inbound conveyor
                       IF  #Cnv_Control.Inputs."Lift Up" THEN
                           #Cnv_Control.Done := FALSE;
                           #Cnv_Control.Instruction.Transfer_in_Progress := TRUE;
                           #Cnv_Control.Current_Task_ID := #Cnv_Control.Instruction.Task_ID;
                           #State := 20;// Roller Running (Popup Up)
                       ELSIF "Pick Station" AND
                           #Cnv_Control.Inputs."Lift Down" (*AND "Control_DB".PopUp_Cnv[4].Inputs."Lift Down"*) THEN //TO pick station
                           #Cnv_Control.Done := FALSE;
                           #Cnv_Control.Instruction.Transfer_in_Progress := TRUE;
                           #Cnv_Control.Current_Task_ID := #Cnv_Control.Instruction.Task_ID;
                           #State := 30;// Chain Running (Popup Down) 
                       ELSIF NOT "Pick Station" (*AND "Control_DB".PopUp_Cnv[4].Inputs."Lift Down"*) THEN //FROM pick station
                           #Cnv_Control.Done := FALSE;
                           #Cnv_Control.Instruction.Transfer_in_Progress := TRUE;
                           #Cnv_Control.Current_Task_ID := #Cnv_Control.Instruction.Task_ID;
                           #State := 40;
                       ELSE
                           #Cnv_Control.Warning := 1; //Cannot transfer from that conveyor
                       END_IF;

                       //Outbound Transfer    
                   ELSIF #Cnv_Control.Instruction.Outbound_Ready AND NOT #Cnv_Control.Running AND #Cnv_Control.Error = 0 THEN
                       //Check transfer ID TO popup cpnveyor 2
                       IF #Cnv_Control.Inputs."Lift Up" AND "Control_DB".PopUp_Cnv[2].Inputs."Lift Up" THEN
                           #Cnv_Control.Done := FALSE;
                           #Cnv_Control.Instruction.Transfer_in_Progress := TRUE;
                           #Cnv_Control.Current_Task_ID := #Cnv_Control.Instruction.Task_ID;
                           #State := 50;
                       ELSE
                           #Cnv_Control.Warning := 1; //Cannot transfer TO that conveyor
                       END_IF;
                   ELSE
                       #Cnv_Control.Warning := 0;// No task that can be started, yet start bit has been made true.
                   END_IF;
               ELSIF #Cnv_Control.Instruction.Start_Transfer AND "Control_DB".VTD_Control.Current_Level <> 0 THEN
                   //Extractor not at the correct level
                   "Set_Bit_F"(Bit := 2,
                               Bit_Value := 1,
                               Var := #Cnv_Control.Cnv_Errors.Error_Word_3);
               END_IF;
               IF #Cnv_Control.Instruction.Lift_Up THEN
                   #Cnv_Control.Done := FALSE;
                   #State := 60; // Lift UP
               ELSIF #Cnv_Control.Instruction.Lift_Down THEN
                   #Cnv_Control.Done := FALSE;
                   #State := 70; // Lift Down
               END_IF;

           20: // Roller Running (Popup Up)
               #Cnv_Control.Running := TRUE;
               #Cnv_Control.Roller_Motor.Forward := TRUE;
               #Cnv_Control.Roller_Motor.Speed := #Cnv_Settings.Roller_Full_Speed;
               #Transfer_Direction := 'Foward';

               IF "R_TRIG_DB_14".Q OR "PopUp Conveyor 2 - Pallet present 3" THEN
                   #Cnv_Control.Done := TRUE;
                   #Cnv_Control.Roller_Motor.Forward := FALSE;
                   #Cnv_Control.Roller_Motor.Reverse := FALSE;
                   #Cnv_Control.Roller_Motor.Speed := 0;
                   #Transfer_Direction := '';
                   #State := 0;
               END_IF;

               //Monitor the transfer progress
               #Timer_Transfer(IN := "Control_DB".Inbound_Cnv.Running,
                               PT := UINT_TO_TIME(#Cnv_Settings.Roller_Transfer_Time) * 1000);
               //If the watchdog bites, kill the process
               IF #Timer_Transfer.Q THEN //14:1 Transfer timed out
                   "Set_Bit_F"(Bit := 3,
                               Bit_Value := 1,
                               Var := #Cnv_Control.Cnv_Errors.Error_Word_2);
               END_IF;

           30: // Chain Running (Popup Down)
               #Cnv_Control.Running := TRUE;
               #Cnv_Control.Chain_Motor.Forward := TRUE;
               #Cnv_Control.Chain_Motor.Speed := #Cnv_Settings.Chain_Full_Speed;
               #Transfer_Direction := 'Foward';

               IF "R_TRIG_DB_14".Q OR NOT "Pick Station" THEN
                   #Cnv_Control.Done := TRUE;
                   #Cnv_Control.Chain_Motor.Forward := FALSE;
                   #Cnv_Control.Chain_Motor.Reverse := FALSE;
                   #Cnv_Control.Chain_Motor.Speed := 0;
                   #Transfer_Direction := '';
                   #State := 0;
               END_IF;

               //Monitor the transfer progress
               #Timer_Transfer(IN := "LighGuard_Cut-Off Path 01",
                               PT := UINT_TO_TIME(#Cnv_Settings.Chain_Transfer_Time) * 1000);
               //If the watchdog bites, kill the process
               IF #Timer_Transfer.Q THEN //14:1 Transfer timed out
                   "Set_Bit_F"(Bit := 3,
                               Bit_Value := 1,
                               Var := #Cnv_Control.Cnv_Errors.Error_Word_2);
               END_IF;

           40: // Chain Running (Popup Down)
               #Cnv_Control.Running := TRUE;
               #Cnv_Control.Chain_Motor.Forward := TRUE;
               #Cnv_Control.Chain_Motor.Speed := #Cnv_Settings.Chain_Full_Speed;
               #Transfer_Direction := 'Foward';

               IF "R_TRIG_DB_14".Q OR "PopUp Conveyor 1 - Pallet sensor" THEN
                   #Cnv_Control.Done := TRUE;
                   #Cnv_Control.Chain_Motor.Forward := FALSE;
                   #Cnv_Control.Chain_Motor.Reverse := FALSE;
                   #Cnv_Control.Chain_Motor.Speed := 0;
                   #Transfer_Direction := '';
                   #State := 0;
               END_IF;

               //Monitor the transfer progress
               #Timer_Transfer(IN := "LighGuard_Cut-Off Path 01",
                               PT := UINT_TO_TIME(#Cnv_Settings.Chain_Transfer_Time) * 1000);
               //If the watchdog bites, kill the process
               IF #Timer_Transfer.Q THEN //14:1 Transfer timed out
                   "Set_Bit_F"(Bit := 3,
                               Bit_Value := 1,
                               Var := #Cnv_Control.Cnv_Errors.Error_Word_2);
               END_IF;

           50: // Roller Running (Popup Up)
               IF "Control_DB".PopUp_Cnv[2].Roller_Motor.Status.%X0 THEN//Is running
                   #Cnv_Control.Running := TRUE;
                   #Cnv_Control.Roller_Motor.Forward := TRUE;
                   #Cnv_Control.Roller_Motor.Speed := #Cnv_Settings.Roller_Full_Speed;
                   #Transfer_Direction := 'Foward';
               END_IF;

               IF "R_TRIG_DB_14".Q OR "PopUp Conveyor 2 - Pallet present 4" THEN
                   #Cnv_Control.Done := TRUE;
                   #Cnv_Control.Roller_Motor.Forward := FALSE;
                   #Cnv_Control.Roller_Motor.Reverse := FALSE;
                   #Cnv_Control.Roller_Motor.Speed := 0;
                   #Transfer_Direction := '';
                   #State := 0;
               END_IF;

               //Monitor the transfer progress
               #Timer_Transfer(IN := TRUE,
                               PT := UINT_TO_TIME(#Cnv_Settings.Roller_Transfer_Time) * 1000);
               //If the watchdog bites, kill the process
               IF #Timer_Transfer.Q THEN //14:1 Transfer timed out
                   "Set_Bit_F"(Bit := 3,
                               Bit_Value := 1,
                               Var := #Cnv_Control.Cnv_Errors.Error_Word_2);
               END_IF;

           60: // Lift Up
               #Cnv_Control.Running := TRUE;
               #Cnv_Control.Lift_Motor.Forward := TRUE;
               #Cnv_Control.Lift_Motor.Speed := #Cnv_Settings.Lift_Full_Speed;
               #Transfer_Direction := 'Up';

               IF #Cnv_Control.Inputs."Lift Up" THEN
                   #Cnv_Control.Done := TRUE;
                   #Cnv_Control.Lift_Motor.Forward := FALSE;
                   #Cnv_Control.Lift_Motor.Reverse := FALSE;
                   #Cnv_Control.Lift_Motor.Speed := 0;
                   #Transfer_Direction := '';
                   #State := 0;
               END_IF;

               //Monitor the transfer progress
               #Timer_Transfer(IN := "LighGuard_Cut-Off Path 01",
                               PT := UINT_TO_TIME(#Cnv_Settings.Lift_Transfer_Time) * 1000);
               //If the watchdog bites, kill the process
               IF #Timer_Transfer.Q THEN //14:1 Transfer timed out
                   "Set_Bit_F"(Bit := 3,
                               Bit_Value := 1,
                               Var := #Cnv_Control.Cnv_Errors.Error_Word_2);
               END_IF;

           70: // Lift Down
               #Cnv_Control.Running := TRUE;
               #Cnv_Control.Lift_Motor.Reverse := TRUE;
               #Cnv_Control.Lift_Motor.Speed := #Cnv_Settings.Lift_Full_Speed;
               #Transfer_Direction := 'Down';

               IF #Cnv_Control.Inputs."Lift Down" THEN
                   #Cnv_Control.Done := TRUE;
                   #Cnv_Control.Lift_Motor.Forward := FALSE;
                   #Cnv_Control.Lift_Motor.Reverse := FALSE;
                   #Cnv_Control.Lift_Motor.Speed := 0;
                   #Transfer_Direction := '';
                   #State := 0;
               END_IF;

               //Monitor the transfer progress
               #Timer_Transfer(IN := "LighGuard_Cut-Off Path 01",
                               PT := UINT_TO_TIME(#Cnv_Settings.Lift_Transfer_Time) * 1000);
               //If the watchdog bites, kill the process
               IF #Timer_Transfer.Q THEN //14:1 Transfer timed out
                   "Set_Bit_F"(Bit := 3,
                               Bit_Value := 1,
                               Var := #Cnv_Control.Cnv_Errors.Error_Word_2);
               END_IF;

           400: //Error state
               #Cnv_Control.Running := FALSE;
               #Cnv_Control.Roller_Motor.Speed := 0;
               #Cnv_Control.Chain_Motor.Speed := 0;
               #Cnv_Control.Lift_Motor.Speed := 0;
               #Cnv_Control.Roller_Motor.Forward := FALSE;
               #Cnv_Control.Chain_Motor.Forward := FALSE;
               #Cnv_Control.Lift_Motor.Forward := FALSE;
               #Cnv_Control.Roller_Motor.Reverse := FALSE;
               #Cnv_Control.Chain_Motor.Reverse := FALSE;
               #Cnv_Control.Lift_Motor.Reverse := FALSE;
               #Cnv_Control.Instruction.Stop := FALSE;
               #Cnv_Control.Instruction.Transfer_in_Progress := FALSE;
               #Watchdog(IN := FALSE,
                         PT := T#0S);
               #Timer_TC(IN := FALSE,
                         PT := T#0S);
               #Timer_Transfer(IN := FALSE,
                               PT := T#0S);
               #IEC_Timer_0_Instance_1(IN := FALSE,
                                       PT := T#0S);
               IF #Cnv_Control.Instruction.Reset THEN
                   #Cnv_Control.Warning := 0;
                   #Cnv_Control.Current_Task_ID := 0;
                   #Cnv_Control.Error := FALSE; //Reset the conveyor

                   #Cnv_Control.Cnv_Errors.Error_Word_1 := 0;
                   #Cnv_Control.Cnv_Errors.Error_Word_2 := 0;
                   #Cnv_Control.Cnv_Errors.Error_Word_3 := 0;
                   #Cnv_Control.Cnv_Errors.Error_Word_4 := 0;
                   #State := 0;
               END_IF;

           500:
               IF #Cnv_Control.Enabled THEN
                   REGION ROLLER
                       IF #Cnv_Control.Inputs."Lift Up" AND NOT #Cnv_Control.Inputs."Lift Down" THEN
                           IF #Cnv_Control.Instruction.Roller_Fwd OR #Cnv_Control.Instruction.Start_Transfer THEN
                               #Cnv_Control.Roller_Motor.Speed := #Cnv_Settings.Roller_Manual_Speed;
                               #Cnv_Control.Roller_Motor.Forward := TRUE;
                               #Cnv_Control.Running := TRUE;
                           ELSIF #Cnv_Control.Instruction.Roller_Bwd OR #Cnv_Control.Instruction.Start_Transfer_Backward THEN
                               #Cnv_Control.Roller_Motor.Speed := #Cnv_Settings.Roller_Manual_Speed;
                               #Cnv_Control.Roller_Motor.Reverse := TRUE;
                               #Cnv_Control.Running := TRUE;
                           ELSE
                               #Cnv_Control.Roller_Motor.Speed := 0;
                               #Cnv_Control.Roller_Motor.Forward := FALSE;
                               #Cnv_Control.Roller_Motor.Reverse := FALSE;
                               #Cnv_Control.Running := FALSE;
                           END_IF;
                       END_IF;
                   END_REGION

                   REGION CHAIN
                       IF NOT #Cnv_Control.Inputs."Lift Up" AND #Cnv_Control.Inputs."Lift Down"
                           AND "Control_DB".PopUp_Cnv[4].Inputs."Lift Down" AND NOT "Control_DB".PopUp_Cnv[4].Inputs."Lift Up" THEN
                           IF #Cnv_Control.Instruction.Chain_Fwd OR #Cnv_Control.Instruction.Start_Transfer THEN
                               #Cnv_Control.Chain_Motor.Speed := #Cnv_Settings.Chain_Manual_Speed;
                               #Cnv_Control.Chain_Motor.Forward := TRUE;
                               #Cnv_Control.Running := TRUE;
                           ELSIF #Cnv_Control.Instruction.Chain_Bwd OR #Cnv_Control.Instruction.Start_Transfer_Backward THEN
                               #Cnv_Control.Chain_Motor.Speed := #Cnv_Settings.Chain_Manual_Speed;
                               #Cnv_Control.Chain_Motor.Reverse := TRUE;
                               #Cnv_Control.Running := TRUE;
                           ELSE
                               #Cnv_Control.Chain_Motor.Speed := 0;
                               #Cnv_Control.Chain_Motor.Forward := FALSE;
                               #Cnv_Control.Chain_Motor.Reverse := FALSE;
                               #Cnv_Control.Running := FALSE;
                           END_IF;
                       END_IF;
                   END_REGION

                   REGION LIFT
                       IF NOT #SinaSpeed_Roller.AxisEnabled AND NOT #SinaSpeed_Chain.AxisEnabled THEN
                           IF #Cnv_Control.Instruction.Lift_Up AND NOT #Cnv_Control.Inputs."Lift Up" THEN
                               #Cnv_Control.Lift_Motor.Speed := #Cnv_Settings.Lift_Manual_Speed;
                               #Cnv_Control.Lift_Motor.Forward := TRUE;
                               #Cnv_Control.Running := TRUE;
                           ELSIF #Cnv_Control.Instruction.Lift_Down AND NOT #Cnv_Control.Inputs."Lift Down" THEN
                               #Cnv_Control.Lift_Motor.Speed := #Cnv_Settings.Lift_Manual_Speed;
                               #Cnv_Control.Lift_Motor.Reverse := TRUE;
                               #Cnv_Control.Running := TRUE;
                           ELSE
                               #Cnv_Control.Lift_Motor.Speed := 0;
                               #Cnv_Control.Lift_Motor.Forward := FALSE;
                               #Cnv_Control.Lift_Motor.Reverse := FALSE;
                               #Cnv_Control.Running := FALSE;
                           END_IF;
                       END_IF;
                   END_REGION
               END_IF;

               IF #Cnv_Control.Mode <> 1 AND #Cnv_Control.Mode <> 5 THEN
                   #State := 0;
               END_IF;
       END_CASE;
   END_REGION



   REGION Cyclic Error Checks
       IF NOT "Main_Safety_RTG1_DB".SAFETY_OK_CAROUSEL THEN //11:1
           "Set_Bit_F"(Bit := 0,
                       Bit_Value := 1,
                       Var := #Cnv_Control.Cnv_Errors.Error_Word_1);
       END_IF;

       // IF #Cnv_Control.Instruction.Stop THEN //11:2
       //     "Set_Bit_F"(Bit := 1,
       //                 Bit_Value := 1,
       //                 Var := #Cnv_Control.Cnv_Errors.Error_Word_1);
       // END_IF;

       IF #Cnv_Control.Roller_Motor.Error OR #Cnv_Control.Chain_Motor.Error OR #Cnv_Control.Lift_Motor.Error THEN
           "Set_Bit_F"(Bit := 0,
                       Bit_Value := 1,
                       Var := #Cnv_Control.Cnv_Errors.Error_Word_4);
       END_IF;

       // Pallet Sensor Checks
       // IF #Cnv_Control.Inputs.Lfwd AND #Cnv_Control.Inputs.Rbwd THEN
       //     #Cnv_Control.Error := TRUE; //15:2 Combination of Cnv_Inputs indicates issue in conveyor
       //     "Set_Bit_F"(Bit := 1,
       //                 Bit_Value := 1,
       //                 Var := #Cnv_Control.Cnv_Errors.Error_Word_4);
       //     #State := 400;
       // IF #Cnv_Control.Inputs.Lfwd AND #Cnv_Control.Inputs.Lpd1 AND #Cnv_Control.Inputs.Rpd1 THEN
       //     #Cnv_Control.Error := TRUE; //15:3 Combination of Cnv_Inputs indicates issue in conveyor
       //     "Set_Bit_F"(Bit := 2,
       //                 Bit_Value := 1,
       //                 Var := #Cnv_Control.Cnv_Errors.Error_Word_4);
       //     #State := 400;
       // ELSIF #Cnv_Control.Inputs.Rbwd AND #Cnv_Control.Inputs.Lpd1 AND #Cnv_Control.Inputs.Rpd1 THEN
       //     #Cnv_Control.Error := TRUE; //15:4 Combination of Cnv_Inputs indicates issue in conveyor
       //     "Set_Bit_F"(Bit := 3,
       //                 Bit_Value := 1,
       //                 Var := #Cnv_Control.Cnv_Errors.Error_Word_4);
       //     #State := 400;
       // END_IF;

       // Shuttle in Place Cnv_Inputs - Need to confirm the order of these Cnv_Inputs.
       // IF (#Cnv_Settings.ID > 110000 AND #Cnv_Settings.ID < 120000 AND NOT #Cnv_Control.Inputs.Sdetect1 AND #Cnv_Control.Inputs.Sdetect2)
       //     OR (#Cnv_Settings.ID > 120000 AND #Cnv_Settings.ID < 130000 AND NOT #Cnv_Control.Inputs.Sdetect1 AND #Cnv_Control.Inputs.Sdetect2) THEN
       //     #Cnv_Control.Error := TRUE; //14:5 Shuttle is about to yeet itself down the VTD shaft
       //     "Set_Bit_F"(Bit := 7,
       //                 Bit_Value := 1,
       //                 Var := #Cnv_Control.Cnv_Errors.Error_Word_2);
       //     #State := 400;
       // END_IF;

       // IF (#Cnv_Settings.ID > 110000 AND #Cnv_Settings.ID < 120000 AND #Cnv_Control.Inputs.Sdetect1 AND NOT #Cnv_Control.Inputs.Sdetect2)
       //     OR (#Cnv_Settings.ID > 120000 AND #Cnv_Settings.ID < 130000 AND #Cnv_Control.Inputs.Sdetect1 AND NOT #Cnv_Control.Inputs.Sdetect2) THEN
       //     #Cnv_Control.Warning := 0; //Shuttle detected in conveyor not yet on barcode
       // END_IF;

       // // #Watchdog auto starts the moment Any form OF transfer occurs.
       // IF #State > 10 AND #State < 400 THEN
       //     #Watchdog(IN := TRUE,
       //               PT := T#200s);
       // ELSE
       //     #Watchdog.IN := FALSE;
       // END_IF;

       // IF #Watchdog.Q THEN
       //     #Watchdog.IN := FALSE;
       //     #Cnv_Control.Error := TRUE; //14:2  Watchdog bit
       //     "Set_Bit_F"(Bit := 4,
       //                 Bit_Value := 1,
       //                 Var := #Cnv_Control.Cnv_Errors.Error_Word_2);
       //     #State := 400;
       // END_IF;

       // go to error state
       IF #Cnv_Control.Cnv_Errors.Error_Word_1 <> 0 OR
           #Cnv_Control.Cnv_Errors.Error_Word_2 <> 0 OR
           #Cnv_Control.Cnv_Errors.Error_Word_3 <> 0 OR
           #Cnv_Control.Cnv_Errors.Error_Word_4 <> 0
       THEN
           #Cnv_Control.Error := TRUE;
           #State := 400;
       END_IF;
   END_REGION

   REGION VFD
       REGION ROLLER
           #Cnv_Control.Roller_Motor.Ready := NOT #Cnv_Control.Roller_Motor.Error;

           #SinaSpeed_Roller(EnableAxis := #Cnv_Control.Roller_Motor.Forward OR #Cnv_Control.Roller_Motor.Reverse,
                             AckError := #Cnv_Control.Instruction.Reset,
                             SpeedSp := #MainSetpoint_Roller,
                             RefSpeed := 1745.0,
                             HWIDSTW := #Cnv_Settings.Roller_G120_Hardware_ID,
                             HWIDZSW := #Cnv_Settings.Roller_G120_Hardware_ID,
                             AxisEnabled => #Cnv_Control.Roller_Motor.Status.%X0,
                             Lockout => #Cnv_Control.Roller_Motor.Error,
                             Error => #Cnv_Control.Roller_Motor.Error);

           //MAIN SETPOINT
           IF #Cnv_Control.Roller_Motor.Reverse THEN
               #MainSetpoint_Roller := (SCALE_X(MIN := 0,
                                                VALUE := NORM_X(MIN := 0,
                                                                VALUE := #Cnv_Control.Roller_Motor.Speed,
                                                                MAX := 100),
                                                MAX := 1745.0) * -1);
           ELSIF #Cnv_Control.Roller_Motor.Forward THEN
               #MainSetpoint_Roller := SCALE_X(MIN := 0,
                                               VALUE := NORM_X(MIN := 0,
                                                               VALUE := #Cnv_Control.Roller_Motor.Speed,
                                                               MAX := 100),
                                               MAX := 1745.0);
           ELSE
               #MainSetpoint_Roller := 0;
           END_IF;

           REGION Actual Speed
               IF #MainSetpoint_Roller > 0 THEN
                   #Cnv_Control.Roller_Motor.Speed_Actual := SCALE_X(MIN := 0,
                                                                     VALUE := NORM_X(MIN := 0,
                                                                                     VALUE := #SinaSpeed_Roller.ActVelocity,
                                                                                     MAX := 1745.0),
                                                                     MAX := 100);
               ELSIF #MainSetpoint_Roller < 0 THEN
                   #Cnv_Control.Roller_Motor.Speed_Actual := SCALE_X(MIN := 0,
                                                                     VALUE := NORM_X(MIN := 0,
                                                                                     VALUE := #SinaSpeed_Roller.ActVelocity * -1,
                                                                                     MAX := 1745.0),
                                                                     MAX := 100);
               ELSE
                   #Cnv_Control.Roller_Motor.Speed_Actual := 0;
               END_IF;
           END_REGION
       END_REGION

       REGION CHAIN
           #Cnv_Control.Chain_Motor.Ready := NOT #Cnv_Control.Chain_Motor.Error;

           #SinaSpeed_Chain(EnableAxis := (#Cnv_Control.Chain_Motor.Forward OR #Cnv_Control.Chain_Motor.Reverse) AND "LighGuard_Cut-Off Path 01",
                            AckError := #Cnv_Control.Instruction.Reset,
                            SpeedSp := #MainSetpoint_Chain,
                            RefSpeed := 1745.0,
                            HWIDSTW := #Cnv_Settings.Chain_G120_Hardware_ID,
                            HWIDZSW := #Cnv_Settings.Chain_G120_Hardware_ID,
                            AxisEnabled => #Cnv_Control.Chain_Motor.Status.%X0,
                            Lockout => #Cnv_Control.Chain_Motor.Error,
                            Error => #Cnv_Control.Chain_Motor.Error);

           //MAIN SETPOINT
           IF #Cnv_Control.Chain_Motor.Reverse AND "LighGuard_Cut-Off Path 01" THEN
               #MainSetpoint_Chain := (SCALE_X(MIN := 0,
                                               VALUE := NORM_X(MIN := 0,
                                                               VALUE := #Cnv_Control.Chain_Motor.Speed,
                                                               MAX := 100),
                                               MAX := 1745.0) * -1);
           ELSIF #Cnv_Control.Chain_Motor.Forward AND "LighGuard_Cut-Off Path 01" THEN
               #MainSetpoint_Chain := SCALE_X(MIN := 0,
                                              VALUE := NORM_X(MIN := 0,
                                                              VALUE := #Cnv_Control.Chain_Motor.Speed,
                                                              MAX := 100),
                                              MAX := 1745.0);
           ELSE
               #MainSetpoint_Chain := 0;
           END_IF;

           REGION Actual Speed
               IF #MainSetpoint_Chain > 0 THEN
                   #Cnv_Control.Chain_Motor.Speed_Actual := SCALE_X(MIN := 0,
                                                                    VALUE := NORM_X(MIN := 0,
                                                                                    VALUE := #SinaSpeed_Chain.ActVelocity,
                                                                                    MAX := 1745.0),
                                                                    MAX := 100);
               ELSIF #MainSetpoint_Chain < 0 THEN
                   #Cnv_Control.Chain_Motor.Speed_Actual := SCALE_X(MIN := 0,
                                                                    VALUE := NORM_X(MIN := 0,
                                                                                    VALUE := #SinaSpeed_Chain.ActVelocity * -1,
                                                                                    MAX := 1745.0),
                                                                    MAX := 100);
               ELSE
                   #Cnv_Control.Chain_Motor.Speed_Actual := 0;
               END_IF;
           END_REGION
       END_REGION

       REGION LIFT
           #Cnv_Control.Lift_Motor.Ready := NOT #Cnv_Control.Lift_Motor.Error;

           #SinaSpeed_Lift(EnableAxis := (#Cnv_Control.Lift_Motor.Forward OR #Cnv_Control.Lift_Motor.Reverse) AND "LighGuard_Cut-Off Path 01",
                           AckError := #Cnv_Control.Instruction.Reset,
                           SpeedSp := #MainSetpoint_Lift,
                           RefSpeed := 1745.0,
                           HWIDSTW := #Cnv_Settings.Lift_G120_Hardware_ID,
                           HWIDZSW := #Cnv_Settings.Lift_G120_Hardware_ID,
                           AxisEnabled => #Cnv_Control.Lift_Motor.Status.%X0,
                           Lockout => #Cnv_Control.Lift_Motor.Error,
                           Error => #Cnv_Control.Lift_Motor.Error);

           //MAIN SETPOINT
           IF #Cnv_Control.Lift_Motor.Reverse AND "LighGuard_Cut-Off Path 01" THEN
               #MainSetpoint_Lift := (SCALE_X(MIN := 0,
                                              VALUE := NORM_X(MIN := 0,
                                                              VALUE := #Cnv_Control.Lift_Motor.Speed,
                                                              MAX := 100),
                                              MAX := 1745.0) * -1);
           ELSIF #Cnv_Control.Lift_Motor.Forward AND "LighGuard_Cut-Off Path 01" THEN
               #MainSetpoint_Lift := SCALE_X(MIN := 0,
                                             VALUE := NORM_X(MIN := 0,
                                                             VALUE := #Cnv_Control.Lift_Motor.Speed,
                                                             MAX := 100),
                                             MAX := 1745.0);
           ELSE
               #MainSetpoint_Lift := 0;
           END_IF;

           REGION Actual Speed
               IF #MainSetpoint_Lift > 0 THEN
                   #Cnv_Control.Lift_Motor.Speed_Actual := SCALE_X(MIN := 0,
                                                                   VALUE := NORM_X(MIN := 0,
                                                                                   VALUE := #SinaSpeed_Lift.ActVelocity,
                                                                                   MAX := 1745.0),
                                                                   MAX := 100);
               ELSIF #MainSetpoint_Lift < 0 THEN
                   #Cnv_Control.Lift_Motor.Speed_Actual := SCALE_X(MIN := 0,
                                                                   VALUE := NORM_X(MIN := 0,
                                                                                   VALUE := #SinaSpeed_Lift.ActVelocity * -1,
                                                                                   MAX := 1745.0),
                                                                   MAX := 100);
               ELSE
                   #Cnv_Control.Lift_Motor.Speed_Actual := 0;
               END_IF;
           END_REGION
       END_REGION
   END_REGION
END_FUNCTION_BLOCK

FUNCTION "ParseShuttle_Status" : "Shuttle_MQTT_Status_Msg"   // FC16, SCL
{ S7_Optimized_Access := 'TRUE' }
VERSION : 0.1
// stored: AutoNumber true, IsIECCheckEnabled false, SetENOAutomatically false, UDAEnableTagReadback false
   VAR_INPUT
      String_1 : String;
      String_2 : String;
      String_3 : String;
      String_4 : String;
      String_5 : String;
      String_6 : String;
   END_VAR
   VAR CONSTANT
      Empty : String;
   END_VAR
BEGIN
   #ParseShuttle_Status.Request_ID := "FindDINTFieldFragmented"(FieldName := 'requestId',
                                                                Str1 := #String_1,
                                                                Str2:=#Empty);
   #ParseShuttle_Status.Position_ID := "FindDINTFieldFragmented"(FieldName := 'positionId',
                                                                 Str1 := #String_1,
                                                                 Str2 := #Empty);
   #ParseShuttle_Status.Destination_ID := "FindDINTFieldFragmented"(FieldName := 'destinationId',
                                                                    Str1 := #String_1,
                                                                    Str2:=#Empty);
   #ParseShuttle_Status.Distance_Remaining := "FindDINTFieldFragmented"(FieldName := 'distanceRemaining',
                                                                        Str1 := #String_1,
                                                                        Str2 := #Empty);
   #ParseShuttle_Status.Position_X := "FindDINTFieldFragmented"(FieldName := 'positionX',
                                                                Str1 := #String_1,
                                                                Str2 := #Empty);
   #ParseShuttle_Status.Position_Y := "FindDINTFieldFragmented"(FieldName := 'positionY',
                                                                Str1 := #String_1,
                                                                Str2 := #Empty);
   #ParseShuttle_Status.Floor := "FindIntField"(FieldName := 'floor',
                                                   JsonStr := #String_1);
   #ParseShuttle_Status.Operation_Mode := "FindStringField"(FieldName := 'operationMode',
                                                            JsonStr := #String_1);
   #ParseShuttle_Status.Operational_State := "FindStringField"(FieldName := 'operationState',
                                                               JsonStr := #String_2);
   #ParseShuttle_Status.Load_State := "FindStringField"(FieldName := 'loadState',
                                                        JsonStr := #String_2);
   #ParseShuttle_Status.Error_Vehicle_1 := INT_TO_UINT("FindINTFieldFragmented"(FieldName := 'errorVehicle1',
                                                                                                                                    Str1 := #String_2,
                                                                                                                                    Str2:=#String_2));
   #ParseShuttle_Status.Error_Vehicle_2 := INT_TO_UINT("FindIntField"(FieldName := 'errorVehicle2',
                                                                                                                          JsonStr := #String_2));
   #ParseShuttle_Status.Error_Vehicle_3 := INT_TO_UINT("FindIntField"(FieldName := 'errorVehicle3',
                                                                                                                          JsonStr := #String_3));
   #ParseShuttle_Status.Error_Vehicle_4 := INT_TO_UINT("FindIntField"(FieldName := 'errorVehicle4',
                                                                                                                          JsonStr := #String_3));
   #ParseShuttle_Status.Error_Vehicle_5 := INT_TO_UINT("FindIntField"(FieldName := 'errorVehicle5',
                                                                                                                          JsonStr := #String_3));
   #ParseShuttle_Status.Error_Vehicle_6 := INT_TO_UINT("FindIntField"(FieldName := 'errorVehicle6',
                                                                                                                          JsonStr := #String_4));
   #ParseShuttle_Status.Sensor_Inputs := INT_TO_UINT("FindIntField"(FieldName := 'sensorInputs',
                                                                                                                      JsonStr := #String_4));
   #ParseShuttle_Status.Sensor_Outputs := INT_TO_UINT("FindIntField"(FieldName := 'sensorOutputs',
                                                                                                                        JsonStr := #String_4));
   #ParseShuttle_Status.Reader_Value := "FindDINTFieldFragmented"(FieldName := 'readerValue',
                                                                  Str1 := #String_4,
                                                                Str2 := #Empty);
   #ParseShuttle_Status.Pallet_Type := "FindStringField"(FieldName := 'palletType',
                                                         JsonStr := #String_4);
   #ParseShuttle_Status.Energy_Level := INT_TO_UINT("FindINTFieldFragmented"(FieldName := 'energyLevel',
                                                                                                                              Str1 := #String_5,
                                                                                                                              Str2:=#String_5));
   #ParseShuttle_Status.Battery_Voltage := INT_TO_UINT("FindIntField"(FieldName := 'batteryVoltage',
                                                                                                                          JsonStr := #String_5));
   #ParseShuttle_Status.Paused := "FindBoolField"(FieldName := 'paused',
                                                  JsonStr := #String_5);
   #ParseShuttle_Status.Last_Received_Order_ID := "FindIntField"(FieldName := 'lastReceivedOrderId',
                                                                 JsonStr := #String_5);
    #ParseShuttle_Status.Current_Order_ID := "FindIntField"(FieldName := 'currentOrderId',
                                                            JsonStr := #String_6);
          #ParseShuttle_Status.Last_Finished_Order_ID := "FindIntField"(FieldName := 'lastFinishedOrderId',
                                                                        JsonStr := #String_6);
END_FUNCTION

FUNCTION "RemovePlusSign" : String   // FC14, SCL
{ S7_Optimized_Access := 'TRUE' }
VERSION : 0.1
// stored: AutoNumber true, IsIECCheckEnabled false, SetENOAutomatically false, UDAEnableTagReadback false
   VAR_INPUT
      inString : String;
   END_VAR
   VAR_TEMP
      tempString : String;
   END_VAR
BEGIN

   IF LEFT(IN := #inString, L := 1) = '+' THEN
       #tempString := RIGHT(IN := #inString, L := LEN(#inString) - 1);
   ELSE
       #tempString := #inString;
   END_IF;

   #RemovePlusSign := #tempString;
END_FUNCTION

FUNCTION_BLOCK "SAI_IND_WriteDigitalOutputs"   // FB3, LAD
{ S7_Optimized_Access := 'FALSE' }
VERSION : 0.1
// stored: AutoNumber true, IsIECCheckEnabled false, SetENOAutomatically false, UDAEnableTagReadback false
   VAR_INPUT
      ID : HW_IO;
      Output1 : Bool;
      Output2 : Bool;
      Output3 : Bool;
      Output4 : Bool;
      Output5 : Bool;
   END_VAR
   VAR_OUTPUT
      Done : Bool;
      Error : Bool;
   END_VAR
   VAR_IN_OUT
      Write : Bool;
   END_VAR
   VAR DB_SPECIFIC
      "Step" : Int;
      Writing : Bool;
      WritePre : Bool;
      BusyNTrig : Bool;
   END_VAR
   VAR
      WRREC { S7_SetPoint := 'True'} : WRREC;
   END_VAR
   VAR_TEMP
      Length : UInt;
   END_VAR
   VAR_TEMP   // added for the SCL form of the ladder/FBD networks
      _w1 : Bool;
      _w2 : Bool;
   END_VAR
BEGIN

REGION Network 1: Initialization
   // Initializes DONE and ERROR output bits
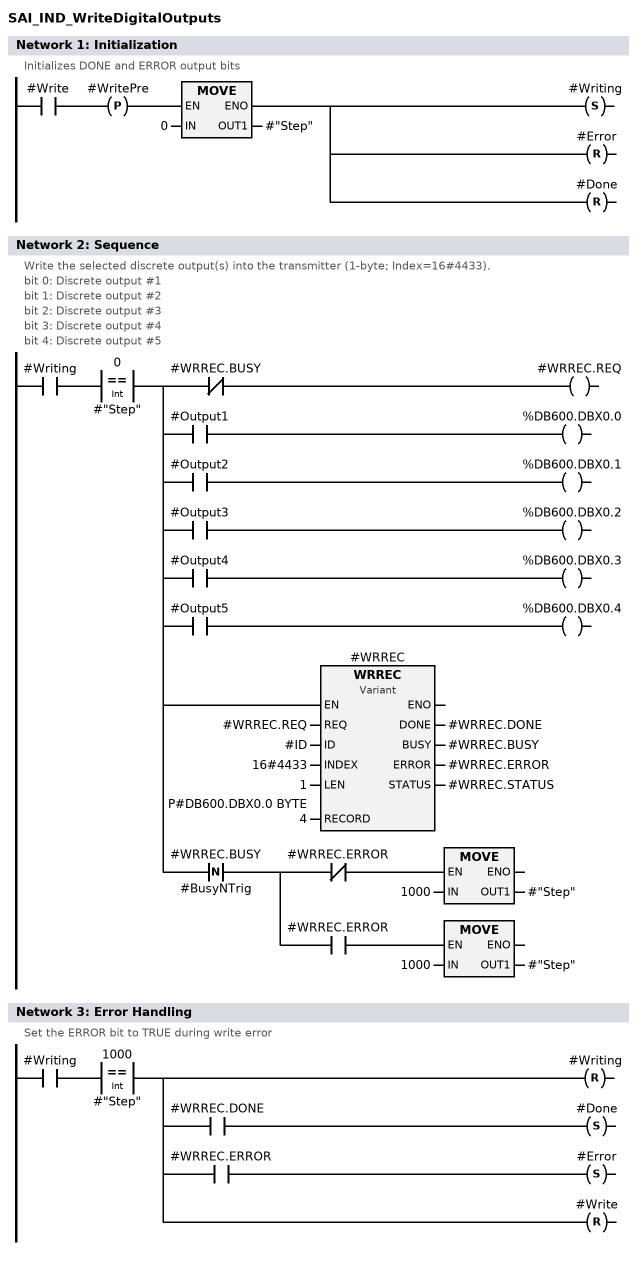
   RUNG wire#powerrail
      Contact( #Write )
      P_Trig( #WritePre )
      { S7_GenerateENO := "TRUE" } Move(in := 0, out1 => #"Step")
      wire#w1
      S_Coil( #Writing )
   END_RUNG
   RUNG wire#w1
      R_Coil( #Error )
   END_RUNG
   RUNG wire#w1
      R_Coil( #Done )
   END_RUNG
   // the same network as SCL:
   // ENO of a box is taken as its EN; it also drops when the box reports an error
   #_w1 := #Write AND NOT #WritePre;   // rising edge
   #WritePre := #Write;
   IF #_w1 THEN
       #"Step" := 0;
       #Writing := TRUE;
       #Error := FALSE;
       #Done := FALSE;
   END_IF;
END_REGION

REGION Network 2: Sequence
   // Write the selected discrete output(s) into the transmitter (1-byte; Index=16#4433).
   // bit 0: Discrete output #1
   // bit 1: Discrete output #2
   // bit 2: Discrete output #3
   // bit 3: Discrete output #4
   // bit 4: Discrete output #5
   RUNG wire#powerrail
      Contact( #Writing )
      { S7_Templates := "SrcType := Int" } EQ_Contact(in1 := 0, in2 := #"Step")
      wire#w1
      I_Contact( #WRREC.BUSY )
      Coil( #WRREC.REQ )
   END_RUNG
   RUNG wire#w1
      Contact( #Output1 )
      Coil( %DB600.DBX0.0 )
   END_RUNG
   RUNG wire#w1
      Contact( #Output2 )
      Coil( %DB600.DBX0.1 )
   END_RUNG
   RUNG wire#w1
      Contact( #Output3 )
      Coil( %DB600.DBX0.2 )
   END_RUNG
   RUNG wire#w1
      Contact( #Output4 )
      Coil( %DB600.DBX0.3 )
   END_RUNG
   RUNG wire#w1
      Contact( #Output5 )
      Coil( %DB600.DBX0.4 )
   END_RUNG
   RUNG wire#w1
      { S7_Templates := "[ptr_type := Variant, id_type := HW_IO, index_type := DInt, len_type := UInt]" } #WRREC.WRREC(REQ := #WRREC.REQ, ID := #ID, INDEX := 16#4433, LEN := 1, RECORD := P#DB600.DBX0.0 BYTE 4, DONE => #WRREC.DONE, BUSY => #WRREC.BUSY, ERROR => #WRREC.ERROR, STATUS => #WRREC.STATUS)
   END_RUNG
   RUNG wire#w1
      N_Contact(operand := #WRREC.BUSY, bit := #BusyNTrig)
      wire#w2
      I_Contact( #WRREC.ERROR )
      { S7_GenerateENO := "TRUE" } Move(in := 1000, out1 => #"Step")
   END_RUNG
   RUNG wire#w2
      Contact( #WRREC.ERROR )
      { S7_GenerateENO := "TRUE" } Move(in := 1000, out1 => #"Step")
   END_RUNG
   // the same network as SCL:
   #_w1 := #Writing AND (0 = #"Step");
   #WRREC.REQ := #_w1 AND NOT #WRREC.BUSY;
   %DB600.DBX0.0 := #_w1 AND #Output1;
   %DB600.DBX0.1 := #_w1 AND #Output2;
   %DB600.DBX0.2 := #_w1 AND #Output3;
   %DB600.DBX0.3 := #_w1 AND #Output4;
   %DB600.DBX0.4 := #_w1 AND #Output5;
   IF #_w1 THEN
       #WRREC(REQ := #WRREC.REQ,   // WRREC
              ID := #ID,
              INDEX := 16#4433,
              LEN := 1,
              RECORD := P#DB600.DBX0.0 BYTE 4,
              DONE => #WRREC.DONE,
              BUSY => #WRREC.BUSY,
              ERROR => #WRREC.ERROR,
              STATUS => #WRREC.STATUS);
   END_IF;
   #_w2 := #_w1 AND NOT #WRREC.BUSY AND #BusyNTrig;   // falling edge of #WRREC.BUSY
   #BusyNTrig := #WRREC.BUSY;
   IF #_w2 AND NOT #WRREC.ERROR THEN #"Step" := 1000; END_IF;
   IF #_w2 AND #WRREC.ERROR THEN #"Step" := 1000; END_IF;
END_REGION

REGION Network 3: Error Handling
   // Set the ERROR bit to TRUE during write error
   RUNG wire#powerrail
      Contact( #Writing )
      { S7_Templates := "SrcType := Int" } EQ_Contact(in1 := 1000, in2 := #"Step")
      wire#w1
      R_Coil( #Writing )
   END_RUNG
   RUNG wire#w1
      Contact( #WRREC.DONE )
      S_Coil( #Done )
   END_RUNG
   RUNG wire#w1
      Contact( #WRREC.ERROR )
      S_Coil( #Error )
   END_RUNG
   RUNG wire#w1
      R_Coil( #Write )
   END_RUNG
   // the same network as SCL:
   #_w1 := #Writing AND (1000 = #"Step");
   IF #_w1 THEN #Writing := FALSE; END_IF;
   IF #_w1 AND #WRREC.DONE THEN #Done := TRUE; END_IF;
   IF #_w1 AND #WRREC.ERROR THEN #Error := TRUE; END_IF;
   IF #_w1 THEN #Write := FALSE; END_IF;
END_REGION
END_FUNCTION_BLOCK

FUNCTION "SICK_GetValue" : Void   // FC10, SCL
TITLE = Get value
{ S7_Optimized_Access := 'TRUE' }
AUTHOR : SICKAG
FAMILY : Ident
VERSION : 1.0
// This function is needs to get a value out of a SICK CoLa command.
// stored: AutoNumber false, IsIECCheckEnabled false, SetENOAutomatically false, UDAEnableTagReadback false
   VAR_INPUT
      iTelegramLength : UInt;   // Length of the source telegram
      iValueLength : USInt;   // ASCII length of the value [1..8] = Fix length | [0]= Variable
      arrData : Array[0..499] of Byte;   // Data record (contains the whole CoLa telegram)
   END_VAR
   VAR_OUTPUT
      nValue : DWord;   // Read value
      nErrorCode : Word;   // Error code
   END_VAR
   VAR_IN_OUT
      iPosition : UInt;   // Position offset of the value before and after (starting from 0)
   END_VAR
   VAR_TEMP
      iLoop : Int;   // Temporarily variable
      iSegmentLength : UInt;   // Length of the segement
      nTemp : DWord;   // Temporarily variable
   END_VAR
BEGIN
   (*===========================================================================================
   Name:   SICK_GetValue
   Author: SICK AG
   =============================================================================================
   Description: 
   This function is for internal use only. The function gets the selected Hex-value string out 
   of the CoLa-Telegram and convert it into a hexadecimal number. 

   =============================================================================================
   Error codes:
   16#0000 = No error
   16#0001 = Invaild telegram length   
   16#0002 = Invalid position index 
   16#0003 = Invalid value length
   16#0004 = Invalid segment length 
   16#0005 = ASCII character is not in a hexadecimal format             

   =============================================================================================
   Version history:
   Date       | Version | created under               | Author  | Remark
   ---------------------------------------------------------------------------------------------
   30/01/2014 | V1.0    | TIA Portal V12 SP1 Update 2 | SICK AG | Initial version
   ============================================================================================*)

   (*===================================== INITIALISATION =====================================*)
   #iSegmentLength:= 0;
   #nValue:= 16#0000_0000;
   #nErrorCode:= 16#0000;

   (*======================================= READ VALUE =======================================*)
   (*Check telegram length*)
   IF #iTelegramLength <=0 OR #iTelegramLength > 500 THEN
     #nErrorCode:= 16#0001; (*Error: Invaild telegram length*)
     RETURN;
   END_IF;

   (*Check current position of the value*)
   IF #iPosition > (#iTelegramLength-1) THEN
     #nErrorCode:= 16#0002; (*Error: Invalid position index*)
     RETURN;
   END_IF;

   (*Check value length*)
   IF #iValueLength >8 THEN
     #nErrorCode:= 16#0003; (*Error: Invalid value length*)
     RETURN;
   END_IF;

   (*Get a value with a variable length (ends with a ' ' or [ETX]*)
   IF #iValueLength = 0 THEN
     FOR #iLoop:= UINT_TO_INT(#iPosition) TO UINT_TO_INT(#iTelegramLength-1) DO
       (*Check if a blank or a [ETX] is detected*)
       IF (#arrData[#iLoop] =' ') OR (#arrData[#iLoop] ='$03') THEN
         EXIT;
       END_IF;

       (*Length of the current value segement*)
       #iSegmentLength:= #iSegmentLength+1;
     END_FOR;

   (*Get a value with a fixed character length [1..8]*)
   ELSE
     #iSegmentLength:= #iValueLength;
   END_IF;

   (*Check if the segment length is valid*)
   IF (#iSegmentLength >8) OR (#iSegmentLength =0) THEN
     #nErrorCode:= 16#0004; (*Error: Invalid segment length*)
     RETURN;
   END_IF;

   (*Convert ASCII string into a hexadecimal number*)
   FOR #iLoop:= UINT_TO_INT(#iPosition) TO UINT_TO_INT(#iPosition+#iSegmentLength-1) DO
     (*ACSII value = [0..9]*)
     IF #arrData[#iLoop] >='0' AND #arrData[#iLoop] <='9' THEN
       #nTemp:= #arrData[#iLoop]-48;
     (*ASCII value = [A..F]*) 
     ELSIF #arrData[#iLoop] >='A' AND #arrData[#iLoop] <='F' THEN
       #nTemp:= #arrData[#iLoop]-55;
     (*ASCII value = [a..f]*)
     ELSIF #arrData[#iLoop] >='a' AND #arrData[#iLoop] <='f' THEN
       #nTemp:= #arrData[#iLoop]-87;    
     ELSE
       #nErrorCode:= 16#0005; (*Error: ASCII character is not in a hexadecimal format *)
       RETURN;
     END_IF;

     (*Create hexadecimal number*)
     #nValue:= SHL(IN:= #nValue, N:= 4);
     #nValue:= #nValue+#nTemp;
   END_FOR;

   (*Set the position of the next element in the telegram*)
   IF #iValueLength = 0 THEN
     #iPosition:= #iPosition+#iSegmentLength+1; (*With blank character*)
   ELSE
     #iPosition:= #iPosition+#iSegmentLength; (*Without blank character*)
   END_IF;
END_FUNCTION

FUNCTION "SICK_SetValue" : Void   // FC11, SCL
TITLE = Set value
{ S7_Optimized_Access := 'TRUE' }
AUTHOR : SICKAG
FAMILY : Ident
VERSION : 1.1
// This function is needs to set a value to a SICK CoLa command.
// stored: AutoNumber false, IsIECCheckEnabled false, SetENOAutomatically false, UDAEnableTagReadback false
   VAR_INPUT
      bAddBlank : Bool;   // Add blank after value
      nValue : DWord;   // Value that should be written
   END_VAR
   VAR_OUTPUT
      arrData : Array[0..499] of Byte;   // Destination telegram
      nErrorCode : Word;   // Error code
   END_VAR
   VAR_IN_OUT
      iPosition : UInt;   // Position offset of the value before and after (starting from 0)
   END_VAR
   VAR_TEMP
      iValueLength : USInt;   // Byte length of the value that shuld be written
      nReturnValue : Word;   // Return value of the convert function
      sValue : String[8];   // Converted value
      nTempValue : DWord;   // Temporarily variable
      iTemp : UInt;   // Temporarily variable
   END_VAR
BEGIN
   (*===========================================================================================
   Name:   SICK_SetValue
   Author: SICK AG
   =============================================================================================
   Description: 
   This function is for internal use only.
   The function converts a hexadecimal value into a hexadecimal string and add it 
   automatically to the command array.     

   =============================================================================================
   Error codes:
   16#0000 = No error
   16#0001 = Invalid position index   
   16#8xxx = Conversion error (HTA-Function) see help system for more information

   =============================================================================================
   Version history:
   Date       | Version | created under               | Author  | Remark
   ---------------------------------------------------------------------------------------------
   30/01/2014 | V1.0    | TIA Portal V12 SP1 Update 2 | SICK AG | Initial version
   22/04/2014 | V1.1    | TIA Portal V12 SP1 Update 4 | SICK AG | Avoid warnings that occur with 
                                                                  TIA V13
   ============================================================================================*)

   (*===================================== INITIALISATION =====================================*)
   #iValueLength:= 0;
   #nErrorCode:= 16#0000;

   (*======================================= WRITE VALUE ======================================*)
   (*Check current position of the value*)
   IF #iPosition > 499 THEN 
     #nErrorCode:= 16#0001; (*Error: Invalid position index*)
     RETURN;
   END_IF;



   (*Get byte length of the value that should be written*)
   IF #nValue <= 16#FF THEN
     #nTempValue:= SHL(IN:= #nValue, N:=24);
     #iValueLength:= 1;
   ELSIF #nValue <= 16#FFFF THEN
     #nTempValue:= SHL(IN:= #nValue, N:=16);
     #iValueLength:= 2;
   ELSIF #nValue <= 16#00FF_FFFF THEN
     #nTempValue:= SHL(IN:= #nValue, N:=8);
     #iValueLength:= 3;
   ELSIF #nValue <= 16#FFFF_FFFF THEN
     #nTempValue:= #nValue;
     #iValueLength:= 4;
   END_IF;

   (*Convert hexadecimal number into a ASCII string*)
   #nReturnValue:= HTA(IN:= #nTempValue, N:= #iValueLength, OUT=>#sValue);
   IF #nReturnValue <> 16#0000 THEN
     #nErrorCode:= #nReturnValue; (*Error: Conversion error (HTA-Function)*)
     RETURN;
   END_IF;

   (*Add the string value to the destination telegram*)
   #arrData[#iPosition]:= 0; // Avoid warnings under TIA V13
   Strg_TO_Chars(Strg:=#sValue, pChars:= #iPosition, Cnt=> #iTemp, Chars:= #arrData);

   (*Add blank to the destination telegram and calculate the position of the next element*)
   IF #bAddBlank THEN
     #arrData[#iPosition+#iTemp]:= ' ';
     #iPosition:= #iPosition+#iTemp+1;

   (*Calculate the position of the next element*)
   ELSE
     #iPosition:= #iPosition+#iTemp;
   END_IF;
END_FUNCTION

FUNCTION "Set_Bit_F" : Void   // FC7, SCL
{ S7_Optimized_Access := 'TRUE' }
VERSION : 0.1
// stored: AutoNumber true, IsIECCheckEnabled false, SetENOAutomatically false, UDAEnableTagReadback false
   VAR_INPUT
      Bit : UInt;
      Bit_Value : Bool;
   END_VAR
   VAR_IN_OUT
      Var : Word;
   END_VAR
BEGIN
   IF #Bit_Value THEN
       // Set the bit
       #Var := #Var OR SHL(IN := WORD#1, N := #Bit);
   // ELSE
   //     // Reset the bit
   //     #Var := #Var OR SHL(IN := DWORD#1, N := #Bit);
   END_IF;
END_FUNCTION

DATA_BLOCK "Barcode_Inbound_FB_DB"   // DB115
VERSION : 0.1
// stored: AutoNumber true, DBAccessibleFromOPCUA true, DBAccessibleFromWebserver true, InstanceOfName Barcode_Station_FB, InstanceOfType FB
"Barcode_Station_FB"
BEGIN
END_DATA_BLOCK

DATA_BLOCK "Barcode_Outbound_FB_DB"   // DB142
VERSION : 0.1
// stored: AutoNumber true, DBAccessibleFromOPCUA true, DBAccessibleFromWebserver true, InstanceOfName Barcode_Station_FB, InstanceOfType FB
"Barcode_Station_FB"
BEGIN
END_DATA_BLOCK

DATA_BLOCK "Barcode_VTD_FB_DB"   // DB144
VERSION : 0.1
// stored: AutoNumber true, DBAccessibleFromOPCUA true, DBAccessibleFromWebserver true, InstanceOfName Barcode_Station_FB, InstanceOfType FB
"Barcode_Station_FB"
BEGIN
END_DATA_BLOCK

DATA_BLOCK "Cnv_L1_FB_DB"   // DB26
AUTHOR : Mertin Coetzee
VERSION : 0.1
// stored: AutoNumber true, DBAccessibleFromOPCUA true, DBAccessibleFromWebserver true, InstanceOfName Buffer_Conveyor_FB, InstanceOfType FB
"Buffer_Conveyor_FB"
BEGIN
END_DATA_BLOCK

DATA_BLOCK "Cnv_L2_FB_DB"   // DB27
AUTHOR : Mertin Coetzee
VERSION : 0.1
// stored: AutoNumber true, DBAccessibleFromOPCUA true, DBAccessibleFromWebserver true, InstanceOfName Buffer_Conveyor_FB, InstanceOfType FB
"Buffer_Conveyor_FB"
BEGIN
END_DATA_BLOCK

DATA_BLOCK "Cnv_L3_FB_DB"   // DB28
AUTHOR : Mertin Coetzee
VERSION : 0.1
// stored: AutoNumber true, DBAccessibleFromOPCUA true, DBAccessibleFromWebserver true, InstanceOfName Buffer_Conveyor_FB, InstanceOfType FB
"Buffer_Conveyor_FB"
BEGIN
END_DATA_BLOCK

DATA_BLOCK "Conveyor_HMI_FB_DB"   // DB73
VERSION : 0.1
// stored: AutoNumber true, DBAccessibleFromOPCUA true, DBAccessibleFromWebserver true, InstanceOfName Conveyor_HMI_FB, InstanceOfType FB
"Conveyor_HMI_FB"
BEGIN
END_DATA_BLOCK

DATA_BLOCK "ECnv_FB_DB"   // DB16
AUTHOR : Mertin Coetzee
VERSION : 0.1
// stored: AutoNumber true, DBAccessibleFromOPCUA true, DBAccessibleFromWebserver true, InstanceOfName EConveyor_FB, InstanceOfType FB
"EConveyor_FB"
BEGIN
END_DATA_BLOCK

DATA_BLOCK "FB_HeartBeat_DB"   // DB136
VERSION : 0.1
// stored: AutoNumber true, DBAccessibleFromOPCUA true, DBAccessibleFromWebserver true, InstanceOfName FB_HeartBeat, InstanceOfType FB
"FB_HeartBeat"
BEGIN
   TimeOut.PT := T#10S;
   TimeOut.IN := TRUE;
   "Timer".PT := T#500MS;
   "Timer".IN := TRUE;
END_DATA_BLOCK

DATA_BLOCK "IDB_SICK_AFx60"   // DB121
VERSION : 0.1
// stored: AutoNumber true, DBAccessibleFromOPCUA true, DBAccessibleFromWebserver true, InstanceOfName FB_SICK_AFx60_PN, InstanceOfType FB
"FB_SICK_AFx60_PN"
BEGIN
END_DATA_BLOCK

DATA_BLOCK "Inbound_Cnv_FB_DB"   // DB30
AUTHOR : Mertin Coetzee
VERSION : 0.1
// stored: AutoNumber true, DBAccessibleFromOPCUA true, DBAccessibleFromWebserver true, InstanceOfName InConveyor_FB, InstanceOfType FB
"InConveyor_FB"
BEGIN
END_DATA_BLOCK

DATA_BLOCK "LCom_Communication_Shuttle1_DB"   // DB65
AUTHOR : APC_ERLF
FAMILY : LCom
VERSION : 2.1
// stored: AutoNumber true, DBAccessibleFromOPCUA true, DBAccessibleFromWebserver true, InstanceOfName LCom_Communication, InstanceOfType FB
"LCom_Communication"
BEGIN
END_DATA_BLOCK

DATA_BLOCK "LCom_Communication_Shuttle2_DB"   // DB67
AUTHOR : APC_ERLF
FAMILY : LCom
VERSION : 2.1
// stored: AutoNumber true, DBAccessibleFromOPCUA true, DBAccessibleFromWebserver true, InstanceOfName LCom_Communication, InstanceOfType FB
"LCom_Communication"
BEGIN
END_DATA_BLOCK

DATA_BLOCK "LCom_Communication_Shuttle3_DB"   // DB79
AUTHOR : APC_ERLF
FAMILY : LCom
VERSION : 2.1
// stored: AutoNumber true, DBAccessibleFromOPCUA true, DBAccessibleFromWebserver true, InstanceOfName LCom_Communication, InstanceOfType FB
"LCom_Communication"
BEGIN
END_DATA_BLOCK

DATA_BLOCK "LMQTT_Client_DB"   // DB18
AUTHOR : Siemens Industry Online Support
FAMILY : LMQTT
VERSION : 4.0
// stored: AutoNumber true, DBAccessibleFromOPCUA true, DBAccessibleFromWebserver true, InstanceOfName LMQTT_Client, InstanceOfType FB
"LMQTT_Client"
BEGIN
END_DATA_BLOCK

DATA_BLOCK "LMQTT_Client_fb"   // DB42
AUTHOR : Siemens Industry Online Support
FAMILY : LMQTT
VERSION : 4.0
// stored: AutoNumber true, DBAccessibleFromOPCUA true, DBAccessibleFromWebserver true, InstanceOfName LMQTT_Client, InstanceOfType FB
"LMQTT_Client"
BEGIN
END_DATA_BLOCK

DATA_BLOCK "LMQTT_DB"   // DB43
{ S7_Optimized_Access := 'TRUE' }
VERSION : 0.1
// stored: AutoNumber true, DBAccessibleFromOPCUA true, DBAccessibleFromWebserver true, InstanceOfName LMQTT_DB_UDT, InstanceOfType UDT, IsOnlyStoredInLoadMemory false, IsWriteProtectedInAS false
"LMQTT_DB_UDT"
   // VAR
   //    enable : Bool;
   //    publish : Bool;
   //    subscribe : Bool;
   //    unsubscribe : Bool;
   //    qos : USInt;
   //    retain : Bool;
   //    publishMsgLen : UDInt;
   //    willMsgLen : UInt;
   //    connParam : "LMQTT_typeConnParam";
   //    clientIdentifier : WString;
   //    username : WString;
   //    password : WString;
   //    willtopic : WString;
   //    willMsgPayload : Array[1..128] of Byte;
   //    mqttTopic : WString;
   //    publishMsgPayload : Array[0..511] of Byte;
   //    receivedTopic : WString;
   //    receivedMsgPayload : Array[0..1024] of Byte;
   //    valid : Bool;
   //    done : Bool;
   //    busy : Bool;
   //    error : Bool;
   //    status : Word;
   //    diagnostics : "typeDiagnostics";
   //    receivedMsgStatus : USInt;
   //    receivedMsgDataLen : UDInt;
   // END_VAR
BEGIN
END_DATA_BLOCK

DATA_BLOCK "Light_Bars_DB"   // DB41
VERSION : 0.1
// stored: AutoNumber true, DBAccessibleFromOPCUA true, DBAccessibleFromWebserver true, InstanceOfName Light_Bars, InstanceOfType FB
"Light_Bars"
BEGIN
END_DATA_BLOCK

DATA_BLOCK "MB_Device_Status"   // DB119
{ S7_Optimized_Access := 'TRUE' }
VERSION : 0.1
// stored: AutoNumber true, DBAccessibleFromOPCUA true, DBAccessibleFromWebserver true, InstanceOfName SAI_MB_DeviceStatus, InstanceOfType UDT, IsOnlyStoredInLoadMemory false, IsWriteProtectedInAS false
"SAI_MB_DeviceStatus"
   // VAR
   //    "Alternate weight unit" : Bool;
   //    "Run flat" : Bool;
   //    "Device specific bit 2" : Bool;
   //    "Device specific bit 3" : Bool;
   //    "Device specific bit 4" : Bool;
   //    "Device specific bit 5" : Bool;
   //    "Device specific bit 6" : Bool;
   //    "Device specific bit 7" : Bool;
   //    "Sequence bit 0" : Bool;
   //    "Sequence bit 1" : Bool;
   //    "Heart Beat" : Bool;
   //    "Data OK" : Bool;
   //    "Alarm Condition" : Bool;
   //    "Center of Zero" : Bool;
   //    Motion : Bool;
   //    "Net Mode" : Bool;
   // END_VAR
BEGIN
END_DATA_BLOCK

DATA_BLOCK "MQTT_Handler_FB_DB"   // DB44
VERSION : 0.1
// stored: AutoNumber true, DBAccessibleFromOPCUA true, DBAccessibleFromWebserver true, InstanceOfName MQTT_Handler_FB, InstanceOfType FB
"MQTT_Handler_FB"
BEGIN
END_DATA_BLOCK

DATA_BLOCK "Main_Safety_RTG1_DB"   // DB1, F_DB
NAME : FUSI
VERSION : 0.1
// stored: AutoNumber true, DBAccessibleFromOPCUA true, DBAccessibleFromWebserver true, InstanceOfName Main_Safety_RTG1, InstanceOfType FB
"Main_Safety_RTG1"
BEGIN
END_DATA_BLOCK

DATA_BLOCK "OPC_UA_Control_FB_DB"   // DB17
VERSION : 0.1
// stored: AutoNumber true, DBAccessibleFromOPCUA true, DBAccessibleFromWebserver true, InstanceOfName OPC_UA_Control_FB, InstanceOfType FB
"OPC_UA_Control_FB"
BEGIN
END_DATA_BLOCK

DATA_BLOCK "Order_Table_FB_Carousel_DB"   // DB138
VERSION : 0.1
// stored: AutoNumber true, DBAccessibleFromOPCUA true, DBAccessibleFromWebserver true, InstanceOfName Order_Table_FB_Carousel, InstanceOfType FB
"Order_Table_FB_Carousel"
BEGIN
END_DATA_BLOCK

DATA_BLOCK "Order_Table_FB_VTD_DB"   // DB139
VERSION : 0.1
// stored: AutoNumber true, DBAccessibleFromOPCUA true, DBAccessibleFromWebserver true, InstanceOfName Order_Table_FB_VTD, InstanceOfType FB
"Order_Table_FB_VTD"
BEGIN
END_DATA_BLOCK

DATA_BLOCK "Outbound_Cnv_FB_DB"   // DB6
AUTHOR : Mertin Coetzee
VERSION : 0.1
// stored: AutoNumber true, DBAccessibleFromOPCUA true, DBAccessibleFromWebserver true, InstanceOfName OutConveyor_FB, InstanceOfType FB
"OutConveyor_FB"
BEGIN
END_DATA_BLOCK

DATA_BLOCK "PConveyor_1_FB_DB"   // DB13
AUTHOR : Mertin Coetzee
VERSION : 0.1
// stored: AutoNumber true, DBAccessibleFromOPCUA true, DBAccessibleFromWebserver true, InstanceOfName PConveyor_1_FB, InstanceOfType FB
"PConveyor_1_FB"
BEGIN
END_DATA_BLOCK

DATA_BLOCK "PConveyor_2_FB_DB"   // DB83
AUTHOR : Mertin Coetzee
VERSION : 0.1
// stored: AutoNumber true, DBAccessibleFromOPCUA true, DBAccessibleFromWebserver true, InstanceOfName PConveyor_2_FB, InstanceOfType FB
"PConveyor_2_FB"
BEGIN
END_DATA_BLOCK

DATA_BLOCK "PConveyor_3_FB_DB"   // DB88
AUTHOR : Mertin Coetzee
VERSION : 0.1
// stored: AutoNumber true, DBAccessibleFromOPCUA true, DBAccessibleFromWebserver true, InstanceOfName PConveyor_3_FB, InstanceOfType FB
"PConveyor_3_FB"
BEGIN
END_DATA_BLOCK

DATA_BLOCK "PConveyor_4_FB_DB"   // DB89
AUTHOR : Mertin Coetzee
VERSION : 0.1
// stored: AutoNumber true, DBAccessibleFromOPCUA true, DBAccessibleFromWebserver true, InstanceOfName PConveyor_4_FB, InstanceOfType FB
"PConveyor_4_FB"
BEGIN
END_DATA_BLOCK

DATA_BLOCK "PickConveyor_FB_DB"   // DB151
AUTHOR : Mertin Coetzee
VERSION : 0.1
// stored: AutoNumber true, DBAccessibleFromOPCUA true, DBAccessibleFromWebserver true, InstanceOfName PickConveyor_FB, InstanceOfType FB
"PickConveyor_FB"
BEGIN
END_DATA_BLOCK

DATA_BLOCK "Profile_Station_DB"   // DB130
{ S7_Optimized_Access := 'TRUE' }
VERSION : 0.1
// stored: AutoNumber true, DBAccessibleFromOPCUA true, DBAccessibleFromWebserver true, InstanceOfName Stations_DB_UDT, InstanceOfType UDT, IsOnlyStoredInLoadMemory false, IsWriteProtectedInAS false
"Stations_DB_UDT"
   // VAR
   //    Enable { ExternalWritable := 'False'} : Bool;
   //    Execute { ExternalWritable := 'False'} : Bool;
   //    Mode : UInt;
   //    Cancel : Bool;
   //    Enabled { ExternalWritable := 'False'} : Bool;
   //    Done { ExternalWritable := 'False'} : Bool;
   //    Running { ExternalWritable := 'False'} : Bool;
   //    CarSize { ExternalWritable := 'False'} : DInt;
   //    strState { ExternalWritable := 'False'} : String;
   // END_VAR
BEGIN
END_DATA_BLOCK

DATA_BLOCK "SAI_Cyclic_CheckAlive_DB"   // DB12
VERSION : 0.1
// stored: AutoNumber true, DBAccessibleFromOPCUA true, DBAccessibleFromWebserver true, InstanceOfName SAI_Cyclic_CheckAlive, InstanceOfType FB
"SAI_Cyclic_CheckAlive"
BEGIN
END_DATA_BLOCK

DATA_BLOCK "SAI_Cyclic_WeightProc_DB"   // DB29
VERSION : 0.1
// stored: AutoNumber true, DBAccessibleFromOPCUA true, DBAccessibleFromWebserver true, InstanceOfName SAI_Cyclic_WeightProc, InstanceOfType FB
"SAI_Cyclic_WeightProc"
BEGIN
END_DATA_BLOCK

DATA_BLOCK "SAI_IND_AlibiRead_DB"   // DB107
VERSION : 0.1
// stored: AutoNumber true, DBAccessibleFromOPCUA true, DBAccessibleFromWebserver true, InstanceOfName SAI_IND360Base_AlibiRead, InstanceOfType FB
"SAI_IND360Base_AlibiRead"
BEGIN
END_DATA_BLOCK

DATA_BLOCK "SAI_IND_CalFree_DB"   // DB112
VERSION : 0.1
// stored: AutoNumber true, DBAccessibleFromOPCUA true, DBAccessibleFromWebserver true, InstanceOfName SAI_IND_CalFree, InstanceOfType FB
"SAI_IND_CalFree"
BEGIN
END_DATA_BLOCK

DATA_BLOCK "SAI_IND_ReadAdjustSettings_DB"   // DB108
VERSION : 0.1
// stored: AutoNumber true, DBAccessibleFromOPCUA true, DBAccessibleFromWebserver true, InstanceOfName SAI_IND_ReadAdjustSettings, InstanceOfType FB
"SAI_IND_ReadAdjustSettings"
BEGIN
END_DATA_BLOCK

DATA_BLOCK "SAI_IND_SpanAdjust_DB"   // DB113
VERSION : 0.1
// stored: AutoNumber true, DBAccessibleFromOPCUA true, DBAccessibleFromWebserver true, InstanceOfName SAI_IND_SpanAdjust, InstanceOfType FB
"SAI_IND_SpanAdjust"
BEGIN
END_DATA_BLOCK

DATA_BLOCK "SAI_IND_WriteAdjustSettings_DB"   // DB109
VERSION : 0.1
// stored: AutoNumber true, DBAccessibleFromOPCUA true, DBAccessibleFromWebserver true, InstanceOfName SAI_IND_WriteAdjustSettings, InstanceOfType FB
"SAI_IND_WriteAdjustSettings"
BEGIN
END_DATA_BLOCK

